        $ 2172 "Weight_value≔get_weight()" "noBreak"
        global Weight_value=get_weight()
        $ 2173 "tilt_angle≔-1" "noBreak"
        global tilt_angle=-1
        $ 2174 "Wait: 0.5" "noBreak"
        sleep(0.5)
        $ 2175 "vib_mot_thread≔ False " "noBreak"
        global vib_mot_thread=  False
        $ 2176 "MoveL" "noBreak"
        $ 2177 "dispense_pos" "noBreak"
        movel(dispense_pos, a=0.2, v=0.05)
        $ 2178 "Integral_error≔0" "noBreak"
        global Integral_error=0
        $ 2179 "current_error≔0" "noBreak"
        global current_error=0
        $ 2180 "previous_error≔0" "noBreak"
        global previous_error=0
        $ 2181 "Set AO[0]=0.0" "noBreak"
        set_standard_analog_out(0, 0.0)
        # begin: URCap Program Node
        #   Source: SensoPart VISOR Robotic, 2.0.0, SensoPart Industriesensorik GmbH
        #   Type: Exit Pose
        $ 2182 "Exit Pose" "noBreak"
        movel(pose_trans(easyPickPose,p[0.0000,0.0000,-0.0000,0.0000,0.0000,0.0000]),a=0.5000,v=0.2500,t=0.000000,r=0.000000)
        # end: URCap Program Node
        easyPickObjTaken = True
      end
      # end: URCap Program Node
      # begin: URCap Program Node
      #   Source: SensoPart VISOR Robotic, 2.0.0, SensoPart Industriesensorik GmbH
      #   Type: No Object Detected
      $ 2183 "No Object Detected" "noBreak"
      if (visor_partsFound(easyPickVisorId) < 1):
        $ 2184 "Popup: No weigh scale detected" "noBreak"
        popup("No weigh scale detected", "Message", False, False, blocking=True)
        else:
      end
      # end: URCap Program Node
    end
    easyPickCount_4 = easyPickCount_4 + 1
    visor_easyPickUpdate(easyPickVisorId, "counter", easyPickCount_4)
    visor_easyPickSetIdent("b1dffd", easyPickVisorId)
    # end: URCap Program Node
  end
  visorFuncEasyPick_a4e600()
  # end: URCap Program Node
  $ 2185 "powder dispensing"
  $ 2187 "Loop Weight_value<Target_weight"
  while (Weight_value<Target_weight):
    $ 2188 "MoveL"
    $ 2189 "Waypoint_75" "breakAfter"
    movel(Waypoint_75_p, a=0.3, v=0.05, r=0.05)
    $ 2190 "ftr_scoop2" "breakAfter"
    movel(ftr_scoop2_p, a=0.3, v=0.05)
    $ 2191 "aftr_scoop1" "breakAfter"
    movel(aftr_scoop1_p, a=0.3, v=0.05)
    $ 2192 "After_disp_3" "breakAfter"
    movel(After_disp_3_p, a=0.3, v=0.05)
    $ 2193 "Loop 1 times"
    Loop_13 = 0
    while (Loop_13 < 1):
      $ 2194 "Waypoint_55" "breakAfter"
      global move_thread_flag_2194=0
      thread move_thread_2194():
        enter_critical
        move_thread_flag_2194 = 1
        movel(Waypoint_55_p, a=0.5, v=0.07)
        move_thread_flag_2194 = 2
        exit_critical
      end
      move_thread_flag_2194 = 0
      move_thread_han_2194 = run move_thread_2194()
      while (True):
        sleep(1.0E-10)
        if (move_thread_flag_2194 > 1):
          join move_thread_han_2194
          break
        end
        sync()
      end
      $ 2196 "Waypoint_56" "breakAfter"
      movel(Waypoint_56_p, a=0.3, v=0.05)
      $ 2197 "Waypoint_74" "breakAfter"
      movel(Waypoint_74_p, a=0.3, v=0.05)
      $ 2198 "Set AO[0]=3.0"
      set_standard_analog_out(0, 0.3)
      $ 2199 "Wait: 2.0"
      sleep(2.0)
      $ 2200 "Set AO[0]=0.0"
      set_standard_analog_out(0, 0.0)
      Loop_13 = Loop_13 + 1
    end
    $ 2201 "ftr_scoop2" "breakAfter"
    movel(ftr_scoop2_p, a=0.3, v=0.05)
    $ 2202 "aftr_scoo3" "breakAfter"
    movel(aftr_scoo3_p, a=0.3, v=0.05)
    $ 2203 "MoveJ"
    $ 2204 "Waypoint_60" "breakAfter"
    movej(get_inverse_kin(Waypoint_60_p, qnear=Waypoint_60_q), a=0.5235987755982988, v=0.3490658503988659, r=0.05)
    $ 2205 "Waypoint_61" "breakAfter"
    movej(get_inverse_kin(Waypoint_61_p, qnear=Waypoint_61_q), a=0.5235987755982988, v=0.3490658503988659, r=0.05)
    $ 2206 "Waypoint_62" "breakAfter"
    movej(get_inverse_kin(Waypoint_62_p, qnear=Waypoint_62_q), a=0.5235987755982988, v=0.3490658503988659)
    $ 2207 "MoveL"
    $ 2208 "Start_thread≔ True "
    global Start_thread=  True
    $ 2209 "dispense_pos" "breakAfter"
    movel(dispense_pos, a=0.2, v=0.05)
    $ 2210 "vib_mot_thread≔ True "
    global vib_mot_thread=  True
    $ 2211 "Wait: 0.5"
    sleep(0.5)
    $ 2212 "Loop Weight_value≤Target_weight and tilt_angle≤-0.40"
    thread Thread_while_2212():
      while (True):
        $ 2213 "current_error≔Target_weight-Weight_value"
        global current_error=Target_weight-Weight_value
        $ 2214 "Integral_error≔Integral_error+current_error*dt"
        global Integral_error=Integral_error+current_error*dt
        $ 2215 "derivative≔(current_error-previous_error)/dt"
        global derivative=(current_error-previous_error)/dt
        $ 2216 "tilt_increment≔(kp*current_error)+(ki*Integral_error)+(kd*derivative)"
        global tilt_increment=(kp*current_error)+(ki*Integral_error)+(kd*derivative)
        $ 2217 "current_pose≔get_actual_tcp_pose()"
        global current_pose= get_actual_tcp_pose ()
        $ 2218 "tilt_angle≔current_pose[4]"
        global tilt_angle=current_pose[4]
        $ 2219 "tilt_pose≔pose_trans(current_pose, p[(tilt_increment/7), 0, 0, 0, tilt_increment, 0])"
        global tilt_pose=pose_trans(current_pose, p[(tilt_increment/7), 0, 0, 0, tilt_increment, 0])
        $ 2220 "movel(tilt_pose, a=0.025, v=0.015, r=0.00001)"
        movel(tilt_pose, a=0.025, v=0.015, r=0.00001)
        $ 2221 "previous_error≔current_error"
        global previous_error=current_error
        $ 2222 "Wait: 0.01"
        sleep(0.01)
      end
    end
    if (Weight_value <= Target_weight  and  tilt_angle <= -0.40):
      global thread_handler_2212=run Thread_while_2212()
      while (Weight_value <= Target_weight  and  tilt_angle <= -0.40):
        sync()
      end
      kill thread_handler_2212
    end
    $ 2223 "Start_thread≔ False "
    global Start_thread=  False
    $ 2224 "Set AO[0]=0.0"
    set_standard_analog_out(0, 0.0)
    $ 2225 "vib_mot_thread≔ False "
    global vib_mot_thread=  False
    $ 2227 "Weight_value≔get_weight()"
    global Weight_value=get_weight()
    $ 2228 "tilt_angle≔-1"
    global tilt_angle=-1
    $ 2229 "Wait: 0.5"
    sleep(0.5)
    $ 2230 "MoveL"
    $ 2231 "dispense_pos" "breakAfter"
    movel(dispense_pos, a=0.2, v=0.05)
    $ 2232 "Integral_error≔0"
    global Integral_error=0
    $ 2233 "current_error≔0"
    global current_error=0
    $ 2234 "previous_error≔0"
    global previous_error=0
  end
  $ 2235 "MoveL"
  $ 2236 "aftr_scoo3" "breakAfter"
  movel(aftr_scoo3_p, a=0.3, v=0.1)
  $ 2237 "ftr_scoop2" "breakAfter"
  movel(ftr_scoop2_p, a=0.4, v=0.1)
  $ 2238 "aftr_scoop1" "breakAfter"
  movel(aftr_scoop1_p, a=0.4, v=0.1)
  $ 2239 "After_disp_3" "breakAfter"
  movel(After_disp_3_p, a=0.4, v=0.1)
  $ 2240 "Set AO[0]=3.0"
  set_standard_analog_out(0, 0.3)
  $ 2241 "Wait: 2.0"
  sleep(2.0)
  $ 2242 "Set AO[0]=0.0"
  set_standard_analog_out(0, 0.0)
  $ 2243 "aftr_scoop1" "breakAfter"
  movel(aftr_scoop1_p, a=1.2, v=0.25)
  $ 2244 "ftr_scoop2" "breakAfter"
  movel(ftr_scoop2_p, a=0.4, v=0.1)
  $ 2245 "Waypoint_63" "breakAfter"
  movel(Waypoint_63_p, a=1.2, v=0.25, r=0.05)
  $ 2246 "Start" "breakAfter"
  movel(Start_p, a=0.6, v=0.15)
  $ 2247 "Popup: Powder dispensed successfully..."
  popup("Powder dispensed successfully...", "Message", False, False, blocking=True)
  elif (38 == switch_1):
    $ 2248 "Case 38"
    $ 2249 "PowderA(M200)"
    # begin: URCap Program Node
    #   Source: SensoPart VISOR Robotic, 2.0.0, SensoPart Industriesensorik GmbH
    #   Type: VISOR Robotic App
    $ 2250 "VISOR Easy Pick"
    def visorFuncEasyPick_cfdeea():
      # begin: URCap Program Node
      #   Source: SensoPart VISOR Robotic, 2.0.0, SensoPart Industriesensorik GmbH
      #   Type: Easy Pick Setup
      $ 2251 "# 1 Setup" "noBreak"
      local easyPickVisorId = 1
      local easyPickArmMounted = True
      local easyPickSetJob = True
      local easyPickJobName = "PowderA"
      local easyPickAtImgAcq = False
      local easyPickImgAcqPose = cont_img_pose
      # end: URCap Program Node
      # begin: URCap Program Node
      #   Source: SensoPart VISOR Robotic, 2.0.0, SensoPart Industriesensorik GmbH
      #   Type: Process
      $ 2252 "Process" "noBreak"
      local easyPickObjTaken = False
      local easyPickTrigger = False
      local easyPickPoseIdx = 0
      local easyPickPose = p[0,0,0,0,0,0]
      def easyPickFuncTrigger(visorId, setJob, jobName, arm):
      if (setJob):
        visor_changeJob(visorId, jobName, 6000)
      end
      if (arm):
        visor_trigger(visorId, 6000, "arm")
      else:
        visor_trigger(visorId, 6000)
      end
      global easyPickParts_6=visor_partsFound(visorId)
      visor_easyPickUpdate(visorId, "parts", visor_partsFound(visorId))
      return visor_getPose3d(visorId, 0)
    end
    while (not easyPickObjTaken):
      easyPickTrigger = (easyPickCount_6 >= visor_partsFound(easyPickVisorId)) or (easyPickCount_6 > 9) or (not visor_easyPickCheckIdent("9c10c0", easyPickVisorId))
      if (easyPickTrigger):
        easyPickCount_6 = 0
      end
      easyPickPoseIdx = easyPickCount_6
      easyPickPose = visor_getPose3d(easyPickVisorId, easyPickPoseIdx)
      visor_easyPickUpdate(easyPickVisorId, "counter", easyPickPoseIdx)
      # begin: URCap Program Node
      #   Source: SensoPart VISOR Robotic, 2.0.0, SensoPart Industriesensorik GmbH
      #   Type: Image Acquisition Pose
      $ 2253 "Image Acquisition Pose" "noBreak"
      if (easyPickTrigger):
        if (not easyPickAtImgAcq):
          movej(pose_trans(easyPickImgAcqPose,p[0.0000,0.0000,-0.0000,0.0000,0.0000,0.0000]),a=1.3963,v=1.0472,t=0.000000,r=0.000000)
          easyPickAtImgAcq = True
        end
        easyPickPose = easyPickFuncTrigger(easyPickVisorId, easyPickSetJob, easyPickJobName, easyPickArmMounted)
      end
      # end: URCap Program Node
      # begin: URCap Program Node
      #   Source: SensoPart VISOR Robotic, 2.0.0, SensoPart Industriesensorik GmbH
      #   Type: Object Detected
      $ 2254 "Object Detected" "noBreak"
      if (visor_partsFound(easyPickVisorId) > 0):
        $ 2255 "Open Gripper" "noBreak"
        # begin: URCap Program Node
        #   Source: Robotiq_Grippers, 1.8.4.4844, Robotiq Inc.
        #   Type: Gripper
        $ 2256 "Gripper Open (1)" "noBreak"
        if not(gripper_connected[0]):
          popup("Gripper 1 must be connected to run this program.", "No connection", False, True, True)
        end
        if not(rq_is_gripper_activated("1")):
          popup("Gripper 1 is not activated. Go to Installation tab > Gripper to activate it and run the program again.", "Not activated", False, True, True)
        end
        rq_set_pos_spd_for(0, 77, 77, "1")
        rq_wait_pos_spe_for_request(0, 77, 77, "1")
        rq_go_to("1")
        rq_wait("1")
        # end: URCap Program Node
        $ 2257 "MoveJ" "noBreak"
        $ 2258 "Waypoint_76" "noBreak"
        movej(get_inverse_kin(Waypoint_76_p, qnear=Waypoint_76_q), a=1.3962634015954636, v=1.0471975511965976)
        # begin: URCap Program Node
        #   Source: SensoPart VISOR Robotic, 2.0.0, SensoPart Industriesensorik GmbH
        #   Type: Approach Pose
        $ 2259 "Approach Pose" "noBreak"
        movej(pose_trans(easyPickPose,p[0.0000,0.0000,0.0500,0.0000,0.0000,0.0000]),a=1.3963,v=1.0472,t=0.000000,r=0.000000)
        # end: URCap Program Node
        # begin: URCap Program Node
        #   Source: SensoPart VISOR Robotic, 2.0.0, SensoPart Industriesensorik GmbH
        #   Type: Target Pose
        $ 2260 "Target Pose" "noBreak"
        movel(pose_trans(easyPickPose,p[0.0000,0.0000,-0.0000,0.0000,0.0000,0.0000]),a=0.5000,v=0.2500,t=0.000000,r=0.000000)
        # end: URCap Program Node
        $ 2261 "Close Gripper" "noBreak"
        # begin: URCap Program Node
        #   Source: Robotiq_Grippers, 1.8.4.4844, Robotiq Inc.
        #   Type: Gripper
        $ 2262 "Gripper Move0mm (1)" "noBreak"
        if not(gripper_connected[0]):
          popup("Gripper 1 must be connected to run this program.", "No connection", False, True, True)
        end
        if not(rq_is_gripper_activated("1")):
          popup("Gripper 1 is not activated. Go to Installation tab > Gripper to activate it and run the program again.", "Not activated", False, True, True)
        end
        rq_set_pos_spd_for(247, 77, 77, "1")
        rq_wait_pos_spe_for_request(247, 77, 77, "1")
        rq_go_to("1")
        rq_wait("1")
        # end: URCap Program Node
        # begin: URCap Program Node
        #   Source: SensoPart VISOR Robotic, 2.0.0, SensoPart Industriesensorik GmbH
        #   Type: Exit Pose
        $ 2263 "Exit Pose" "noBreak"
        movel(pose_trans(easyPickPose,p[0.0000,0.0000,0.0500,0.0000,0.0000,0.0000]),a=0.5000,v=0.2500,t=0.000000,r=0.000000)
        # end: URCap Program Node
        easyPickObjTaken = True
      end
      # end: URCap Program Node
      # begin: URCap Program Node
      #   Source: SensoPart VISOR Robotic, 2.0.0, SensoPart Industriesensorik GmbH
      #   Type: No Object Detected
      $ 2264 "No Object Detected" "noBreak"
      if (visor_partsFound(easyPickVisorId) < 1):
        $ 2265 "Popup: No Powder container is detected" "noBreak"
        popup("No Powder container is detected", "Message", False, False, blocking=True)
        else:
      end
      # end: URCap Program Node
    end
    easyPickCount_6 = easyPickCount_6 + 1
    visor_easyPickUpdate(easyPickVisorId, "counter", easyPickCount_6)
    visor_easyPickSetIdent("9c10c0", easyPickVisorId)
    # end: URCap Program Node
  end
  visorFuncEasyPick_cfdeea()
  # end: URCap Program Node
  $ 2266 "MoveJ"
  $ 2267 "PowderA_wayp1" "breakAfter"
  movej(get_inverse_kin(PowderA_wayp1_p, qnear=PowderA_wayp1_q), a=1.3962634015954636, v=1.0471975511965976, r=0.05)
  $ 2268 "MoveL"
  $ 2269 "Waypoint_80" "breakAfter"
  movel(Waypoint_80_p, a=1.2, v=0.25)
  $ 2270 "MoveL"
  $ 2271 "Decapp_above" "breakAfter"
  movel(Decapp_above_p, a=1.2, v=0.25)
  $ 2272 "Set GRP_3F_Open=On"
  set_standard_digital_out(5, True)
  $ 2273 "Wait: 0.5"
  sleep(0.5)
  $ 2274 "Decapp_place" "breakAfter"
  movel(Decapp_place_p, a=0.3, v=0.05)
  $ 2275 "Set GRP_3F_Open=Off"
  set_standard_digital_out(5, False)
  $ 2276 "Wait: 0.5"
  sleep(0.5)
  # begin: URCap Program Node
  #   Source: Robotiq_Grippers, 1.8.4.4844, Robotiq Inc.
  #   Type: Gripper
  $ 2277 "Gripper Move40mm (1)"
  if not(gripper_connected[0]):
    popup("Gripper 1 must be connected to run this program.", "No connection", False, True, True)
  end
  if not(rq_is_gripper_activated("1")):
    popup("Gripper 1 is not activated. Go to Installation tab > Gripper to activate it and run the program again.", "Not activated", False, True, True)
  end
  rq_set_pos_spd_for(64, 77, 77, "1")
  rq_wait_pos_spe_for_request(64, 77, 77, "1")
  rq_go_to("1")
  rq_wait("1")
  # end: URCap Program Node
  $ 2278 "MoveL"
  $ 2279 "Decapp_above" "breakAfter"
  movel(Decapp_above_p, a=1.2, v=0.25)
  $ 2280 "Waypoint_78" "breakAfter"
  movel(Waypoint_78_p, a=1.2, v=0.25, r=0.05)
  $ 2281 "Home (Safe)"
  movej([-1.2302089344500047, -1.2969853503591224, -1.875639182904262, -1.539621866126728, 1.5731943360401213, -2.80099559440227], a=1.3962634015954636, v=1.0471975511965976)
  elif (39 == switch_1):
    $ 2282 "Case 39"
    $ 2283 "Decap Container A"
    $ 2284 "MoveL"
    $ 2285 "Waypoint_81" "breakAfter"
    movel(Waypoint_81_p, a=1.2, v=0.25)
    $ 2286 "Waypoint_79" "breakAfter"
    movel(Waypoint_79_p, a=1.2, v=0.25)
    # begin: URCap Program Node
    #   Source: Robotiq_Grippers, 1.8.4.4844, Robotiq Inc.
    #   Type: Gripper
    $ 2287 "Gripper Move22mm (1)"
    if not(gripper_connected[0]):
      popup("Gripper 1 must be connected to run this program.", "No connection", False, True, True)
    end
    if not(rq_is_gripper_activated("1")):
      popup("Gripper 1 is not activated. Go to Installation tab > Gripper to activate it and run the program again.", "Not activated", False, True, True)
    end
    rq_set_pos_spd_for(145, 77, 77, "1")
    rq_wait_pos_spe_for_request(145, 77, 77, "1")
    rq_go_to("1")
    rq_wait("1")
    # end: URCap Program Node
    $ 2288 "Decap"
    $ 2289 "Action_Info≔'decapping'"
    global Action_Info="decapping"
    $ 2290 "Set GRP_3F_Enable=On"
    set_standard_digital_out(4, True)
    $ 2291 "Set GRP_3F_Decap=On"
    set_standard_digital_out(3, True)
    $ 2292 "Force"
    sleep(0.02)
    zero_ftsensor()
    force_mode(p[0.0,0.0,0.0,0.0,0.0,0.0], [0, 0, 1, 0, 0, 0], [0.0, 0.0, 2.0, 0.0, 0.0, 0.0], 2, [0.1, 0.1, 5.0E-4, 0.3490658503988659, 0.3490658503988659, 0.3490658503988659])
    $ 2293 "check_decapping(offset=0.010, timeout=4, abort=CMD_Hold)" "noBreak"
    check_decapping(offset=0.010, timeout=4, abort=CMD_Hold)
    end_force_mode()
    stopl(5.0)
    $ 2294 "Set GRP_3F_Decap=Off"
    set_standard_digital_out(3, False)
    $ 2295 "Set GRP_3F_Enable=Off"
    set_standard_digital_out(4, False)
    $ 2296 "MoveL"
    $ 2297 "Waypoint_82" "breakAfter"
    movel(Waypoint_82_p, a=1.2, v=0.25)
    $ 2298 "Cap_above" "breakAfter"
    movel(Cap_above_p, a=1.2, v=0.25, r=0.05)
    $ 2299 "Cap_Place" "breakAfter"
    movel(Cap_Place_p, a=1.2, v=0.25)
    # begin: URCap Program Node
    #   Source: Robotiq_Grippers, 1.8.4.4844, Robotiq Inc.
    #   Type: Gripper
    $ 2300 "Gripper Move39mm (1)"
    if not(gripper_connected[0]):
      popup("Gripper 1 must be connected to run this program.", "No connection", False, True, True)
    end
    if not(rq_is_gripper_activated("1")):
      popup("Gripper 1 is not activated. Go to Installation tab > Gripper to activate it and run the program again.", "Not activated", False, True, True)
    end
    rq_set_pos_spd_for(67, 77, 77, "1")
    rq_wait_pos_spe_for_request(67, 77, 77, "1")
    rq_go_to("1")
    rq_wait("1")
    # end: URCap Program Node
    $ 2301 "Cap_above" "breakAfter"
    movel(Cap_above_p, a=1.2, v=0.25)
    $ 2302 "Home (Safe)"
    movej([-1.2302089344500047, -1.2969853503591224, -1.875639182904262, -1.539621866126728, 1.5731943360401213, -2.80099559440227], a=1.3962634015954636, v=1.0471975511965976)
  elif (40 == switch_1):
    $ 2338 "Case 40"
    $ 2339 "Place the open PowderA container & dosing"
    # begin: URCap Program Node
    #   Source: SensoPart VISOR Robotic, 2.0.0, SensoPart Industriesensorik GmbH
    #   Type: VISOR Robotic App
    $ 2342 "VISOR Easy Pick"
    def visorFuncEasyPick_303fc5():
      # begin: URCap Program Node
      #   Source: SensoPart VISOR Robotic, 2.0.0, SensoPart Industriesensorik GmbH
      #   Type: Easy Pick Setup
      $ 2343 "# 1 Setup" "noBreak"
      local easyPickVisorId = 1
      local easyPickArmMounted = True
      local easyPickSetJob = True
      local easyPickJobName = "PoTS"
      local easyPickAtImgAcq = False
      local easyPickImgAcqPose = cont_img_pose
      # end: URCap Program Node
      # begin: URCap Program Node
      #   Source: SensoPart VISOR Robotic, 2.0.0, SensoPart Industriesensorik GmbH
      #   Type: Process
      $ 2344 "Process" "noBreak"
      local easyPickObjTaken = False
      local easyPickTrigger = False
      local easyPickPoseIdx = 0
      local easyPickPose = p[0,0,0,0,0,0]
      def easyPickFuncTrigger(visorId, setJob, jobName, arm):
      if (setJob):
        visor_changeJob(visorId, jobName, 6000)
      end
      if (arm):
        visor_trigger(visorId, 6000, "arm")
      else:
        visor_trigger(visorId, 6000)
      end
      global easyPickParts_7=visor_partsFound(visorId)
      visor_easyPickUpdate(visorId, "parts", visor_partsFound(visorId))
      return visor_getPose3d(visorId, 0)
    end
    while (not easyPickObjTaken):
      easyPickTrigger = (easyPickCount_7 >= visor_partsFound(easyPickVisorId)) or (easyPickCount_7 > 9) or (not visor_easyPickCheckIdent("2f5077", easyPickVisorId))
      if (easyPickTrigger):
        easyPickCount_7 = 0
      end
      easyPickPoseIdx = easyPickCount_7
      easyPickPose = visor_getPose3d(easyPickVisorId, easyPickPoseIdx)
      visor_easyPickUpdate(easyPickVisorId, "counter", easyPickPoseIdx)
      # begin: URCap Program Node
      #   Source: SensoPart VISOR Robotic, 2.0.0, SensoPart Industriesensorik GmbH
      #   Type: Image Acquisition Pose
      $ 2345 "Image Acquisition Pose" "noBreak"
      if (easyPickTrigger):
        if (not easyPickAtImgAcq):
          movej(pose_trans(easyPickImgAcqPose,p[0.0000,0.0000,-0.0000,0.0000,0.0000,0.0000]),a=1.3963,v=1.0472,t=0.000000,r=0.000000)
          easyPickAtImgAcq = True
        end
        easyPickPose = easyPickFuncTrigger(easyPickVisorId, easyPickSetJob, easyPickJobName, easyPickArmMounted)
      end
      # end: URCap Program Node
      # begin: URCap Program Node
      #   Source: SensoPart VISOR Robotic, 2.0.0, SensoPart Industriesensorik GmbH
      #   Type: Object Detected
      $ 2346 "Object Detected" "noBreak"
      if (visor_partsFound(easyPickVisorId) > 0):
        $ 2347 "Open Gripper" "noBreak"
        # begin: URCap Program Node
        #   Source: Robotiq_Grippers, 1.8.4.4844, Robotiq Inc.
        #   Type: Gripper
        $ 2348 "Gripper Open (1)" "noBreak"
        if not(gripper_connected[0]):
          popup("Gripper 1 must be connected to run this program.", "No connection", False, True, True)
        end
        if not(rq_is_gripper_activated("1")):
          popup("Gripper 1 is not activated. Go to Installation tab > Gripper to activate it and run the program again.", "Not activated", False, True, True)
        end
        rq_set_pos_spd_for(0, 77, 77, "1")
        rq_wait_pos_spe_for_request(0, 77, 77, "1")
        rq_go_to("1")
        rq_wait("1")
        # end: URCap Program Node
        $ 2349 "MoveL" "noBreak"
        $ 2350 "OP_PowderA2" "noBreak"
        movel(OP_PowderA2_p, a=1.2, v=0.25)
        $ 2351 "OP_PowderA_abov" "noBreak"
        movel(OP_PowderA_abov_p, a=1.2, v=0.25)
        $ 2352 "OP_PowderA_pick" "noBreak"
        movel(OP_PowderA_pick_p, a=1.2, v=0.25)
        # begin: URCap Program Node
        #   Source: Robotiq_Grippers, 1.8.4.4844, Robotiq Inc.
        #   Type: Gripper
        $ 2353 "Gripper Close (1)" "noBreak"
        if not(gripper_connected[0]):
          popup("Gripper 1 must be connected to run this program.", "No connection", False, True, True)
        end
        if not(rq_is_gripper_activated("1")):
          popup("Gripper 1 is not activated. Go to Installation tab > Gripper to activate it and run the program again.", "Not activated", False, True, True)
        end
        rq_set_pos_spd_for(255, 77, 77, "1")
        rq_wait_pos_spe_for_request(255, 77, 77, "1")
        rq_go_to("1")
        rq_wait("1")
        # end: URCap Program Node
        $ 2354 "Wait: 0.5" "noBreak"
        sleep(0.5)
        $ 2355 "Set GRP_3F_Open=On" "noBreak"
        set_standard_digital_out(5, True)
        $ 2357 "OP_PowderA_abov" "noBreak"
        movel(OP_PowderA_abov_p, a=0.3, v=0.05)
        $ 2358 "Op_PowA_wP" "noBreak"
        movel(Op_PowA_wP_p, a=1.2, v=0.25)
        # begin: URCap Program Node
        #   Source: SensoPart VISOR Robotic, 2.0.0, SensoPart Industriesensorik GmbH
        #   Type: Approach Pose
        $ 2359 "Approach Pose" "noBreak"
        movej(pose_trans(easyPickPose,p[0.0000,0.0000,-0.0000,0.0000,0.0000,0.0000]),a=0.5236,v=0.4363,t=0.000000,r=0.000000)
        # end: URCap Program Node
        # begin: URCap Program Node
        #   Source: SensoPart VISOR Robotic, 2.0.0, SensoPart Industriesensorik GmbH
        #   Type: Target Pose
        $ 2360 "Target Pose" "noBreak"
        movel(pose_trans(easyPickPose,p[0.0000,0.0000,-0.0000,0.0000,0.0000,0.0000]),a=0.1000,v=0.0500,t=0.000000,r=0.000000)
        # end: URCap Program Node
        $ 2361 "Close Gripper" "noBreak"
        $ 2362 "target_pose≔pose_add(get_actual_tcp_pose(), p[0,0,-0.085,0,0,0])" "noBreak"
        global target_pose=pose_add(get_actual_tcp_pose(), p[0,0,-0.085,0,0,0])
        $ 2363 "MoveL" "noBreak"
        $ 2364 "target_pose" "noBreak"
        movel(target_pose, a=0.3, v=0.05)
        # begin: URCap Program Node
        #   Source: Robotiq_Grippers, 1.8.4.4844, Robotiq Inc.
        #   Type: Gripper
        $ 2365 "Gripper Open (1)" "noBreak"
        if not(gripper_connected[0]):
          popup("Gripper 1 must be connected to run this program.", "No connection", False, True, True)
        end
        if not(rq_is_gripper_activated("1")):
          popup("Gripper 1 is not activated. Go to Installation tab > Gripper to activate it and run the program again.", "Not activated", False, True, True)
        end
        rq_set_pos_spd_for(0, 77, 77, "1")
        rq_wait_pos_spe_for_request(0, 77, 77, "1")
        rq_go_to("1")
        rq_wait("1")
        # end: URCap Program Node
        # begin: URCap Program Node
        #   Source: SensoPart VISOR Robotic, 2.0.0, SensoPart Industriesensorik GmbH
        #   Type: Exit Pose
        $ 2366 "Exit Pose" "noBreak"
        movel(pose_trans(easyPickPose,p[0.0000,0.0000,-0.0000,0.0000,0.0000,0.0000]),a=0.5000,v=0.2500,t=0.000000,r=0.000000)
        # end: URCap Program Node
        easyPickObjTaken = True
      end
      # end: URCap Program Node
      # begin: URCap Program Node
      #   Source: SensoPart VISOR Robotic, 2.0.0, SensoPart Industriesensorik GmbH
      #   Type: No Object Detected
      $ 2367 "No Object Detected" "noBreak"
      if (visor_partsFound(easyPickVisorId) < 1):
        $ 2368 "Popup: No weigh scale detected" "noBreak"
        popup("No weigh scale detected", "Message", False, False, blocking=True)
        else:
      end
      # end: URCap Program Node
    end
    easyPickCount_7 = easyPickCount_7 + 1
    visor_easyPickUpdate(easyPickVisorId, "counter", easyPickCount_7)
    visor_easyPickSetIdent("2f5077", easyPickVisorId)
    # end: URCap Program Node
  end
  visorFuncEasyPick_303fc5()
  # end: URCap Program Node
  $ 2369 "place_pose≔get_actual_tcp_pose()"
  global place_pose= get_actual_tcp_pose ()
  $ 2370 "center_pose()"
  center_pose()
  $ 2371 "center_pose_t≔P_center"
  global center_pose_t=P_center
  $ 2372 "MoveJ"
  $ 2373 "Waypoint_1" "breakAfter"
  movej(get_inverse_kin(Waypoint_1_p, qnear=Waypoint_1_q), a=1.3962634015954636, v=1.0471975511965976)
  elif (41 == switch_1):
    $ 2374 "Case 41"
    $ 2375 "Powder Emptying"
    $ 2376 "zero_scale()"
    zero_scale()
    $ 2377 "Task≔'Emptying'"
    global Task="Emptying"
    # begin: URCap Program Node
    #   Source: SensoPart VISOR Robotic, 2.0.0, SensoPart Industriesensorik GmbH
    #   Type: VISOR Robotic App
    $ 2378 "VISOR Easy Pick"
    def visorFuncEasyPick_221058():
      # begin: URCap Program Node
      #   Source: SensoPart VISOR Robotic, 2.0.0, SensoPart Industriesensorik GmbH
      #   Type: Easy Pick Setup
      $ 2379 "# 1 Setup" "noBreak"
      local easyPickVisorId = 1
      local easyPickArmMounted = True
      local easyPickSetJob = True
      local easyPickJobName = "Weigh_target"
      local easyPickAtImgAcq = False
      local easyPickImgAcqPose = FRM_Weigh_scale
      # end: URCap Program Node
      # begin: URCap Program Node
      #   Source: SensoPart VISOR Robotic, 2.0.0, SensoPart Industriesensorik GmbH
      #   Type: Process
      $ 2380 "Process" "noBreak"
      local easyPickObjTaken = False
      local easyPickTrigger = False
      local easyPickPoseIdx = 0
      local easyPickPose = p[0,0,0,0,0,0]
      def easyPickFuncTrigger(visorId, setJob, jobName, arm):
      if (setJob):
        visor_changeJob(visorId, jobName, 6000)
      end
      if (arm):
        visor_trigger(visorId, 6000, "arm")
      else:
        visor_trigger(visorId, 6000)
      end
      global easyPickParts_4=visor_partsFound(visorId)
      visor_easyPickUpdate(visorId, "parts", visor_partsFound(visorId))
      return visor_getPose3d(visorId, 0)
    end
    while (not easyPickObjTaken):
      easyPickTrigger = (easyPickCount_4 >= visor_partsFound(easyPickVisorId)) or (easyPickCount_4 > 9) or (not visor_easyPickCheckIdent("7aa8bf", easyPickVisorId))
      if (easyPickTrigger):
        easyPickCount_4 = 0
      end
      easyPickPoseIdx = easyPickCount_4
      easyPickPose = visor_getPose3d(easyPickVisorId, easyPickPoseIdx)
      visor_easyPickUpdate(easyPickVisorId, "counter", easyPickPoseIdx)
      # begin: URCap Program Node
      #   Source: SensoPart VISOR Robotic, 2.0.0, SensoPart Industriesensorik GmbH
      #   Type: Image Acquisition Pose
      $ 2381 "Image Acquisition Pose" "noBreak"
      if (easyPickTrigger):
        if (not easyPickAtImgAcq):
          movej(pose_trans(easyPickImgAcqPose,p[0.0000,0.0000,-0.0000,0.0000,0.0000,0.0000]),a=1.3963,v=1.0472,t=0.000000,r=0.000000)
          easyPickAtImgAcq = True
        end
        easyPickPose = easyPickFuncTrigger(easyPickVisorId, easyPickSetJob, easyPickJobName, easyPickArmMounted)
      end
      # end: URCap Program Node
      # begin: URCap Program Node
      #   Source: SensoPart VISOR Robotic, 2.0.0, SensoPart Industriesensorik GmbH
      #   Type: Object Detected
      $ 2382 "Object Detected" "noBreak"
      if (visor_partsFound(easyPickVisorId) > 0):
        $ 2383 "Open Gripper" "noBreak"
        $ 2384 "tare_scale()" "noBreak"
        tare_scale()
        $ 2385 "Wait: 0.2" "noBreak"
        sleep(0.2)
        $ 2386 "Weight_value≔get_weight()" "noBreak"
        global Weight_value=get_weight()
        $ 2387 "Wait: 0.2" "noBreak"
        sleep(0.2)
        $ 2388 "compute_level_percent(W_now, Weight_value)" "noBreak"
        compute_level_percent(W_now, Weight_value)
        $ 2389 "If level≥10.0" "noBreak"
        if (level >= 10.0):
          $ 2390 "MoveJ" "noBreak"
          $ 2391 "Spatula_otw" "noBreak"
          movej(get_inverse_kin(Spatula_otw_p, qnear=Spatula_otw_q), a=1.3962634015954636, v=1.0471975511965976)
          $ 2392 "pick_spat_L_abv" "noBreak"
          movej(get_inverse_kin(pick_spat_L_abv_p, qnear=pick_spat_L_abv_q), a=1.3962634015954636, v=1.0471975511965976)
          $ 2393 "MoveL" "noBreak"
          $ 2394 "spat_L_pick" "noBreak"
          movel(spat_L_pick_p, a=1.2, v=0.25)
          # begin: URCap Program Node
          #   Source: Robotiq_Grippers, 1.8.4.4844, Robotiq Inc.
          #   Type: Gripper
          $ 2395 "Gripper Close (1)" "noBreak"
          if not(gripper_connected[0]):
            popup("Gripper 1 must be connected to run this program.", "No connection", False, True, True)
          end
          if not(rq_is_gripper_activated("1")):
            popup("Gripper 1 is not activated. Go to Installation tab > Gripper to activate it and run the program again.", "Not activated", False, True, True)
          end
          rq_set_pos_spd_for(255, 0, 77, "1")
          rq_wait_pos_spe_for_request(255, 0, 77, "1")
          rq_go_to("1")
          rq_wait("1")
          # end: URCap Program Node
          $ 2396 "spat_L_lift" "noBreak"
          movel(spat_L_lift_p, a=1.2, v=0.25)
          $ 2397 "spat_L_side" "noBreak"
          movel(spat_L_side_p, a=1.2, v=0.25)
          $ 2398 "spat_L_up" "noBreak"
          movel(spat_L_up_p, a=1.2, v=0.25)
          $ 2399 "MoveJ" "noBreak"
          $ 2400 "Spatula_otw" "noBreak"
          movej(get_inverse_kin(Spatula_otw_p, qnear=Spatula_otw_q), a=1.3962634015954636, v=1.0471975511965976)
        else:
          $ 2401 "ElseIf level≥1.0  and level<10.0" "noBreak"
          if (level >= 1.0   and  level<10.0):
            $ 2402 "MoveJ" "noBreak"
            $ 2403 "Spatula_otw" "noBreak"
            movej(get_inverse_kin(Spatula_otw_p, qnear=Spatula_otw_q), a=1.3962634015954636, v=1.0471975511965976)
            $ 2404 "spat_M_up" "noBreak"
            movej(get_inverse_kin(spat_M_up_p, qnear=spat_M_up_q), a=1.3962634015954636, v=1.0471975511965976)
            $ 2405 "MoveL" "noBreak"
            $ 2406 "spat_M_pick" "noBreak"
            movel(spat_M_pick_p, a=1.2, v=0.25)
            # begin: URCap Program Node
            #   Source: Robotiq_Grippers, 1.8.4.4844, Robotiq Inc.
            #   Type: Gripper
            $ 2407 "Gripper Close (1)" "noBreak"
            if not(gripper_connected[0]):
              popup("Gripper 1 must be connected to run this program.", "No connection", False, True, True)
            end
            if not(rq_is_gripper_activated("1")):
              popup("Gripper 1 is not activated. Go to Installation tab > Gripper to activate it and run the program again.", "Not activated", False, True, True)
            end
            rq_set_pos_spd_for(255, 0, 77, "1")
            rq_wait_pos_spe_for_request(255, 0, 77, "1")
            rq_go_to("1")
            rq_wait("1")
            # end: URCap Program Node
            $ 2408 "spat_M_up" "noBreak"
            movel(spat_M_up_p, a=1.2, v=0.25)
            $ 2409 "Spatula_otw" "noBreak"
            movel(Spatula_otw_p, a=1.2, v=0.25)
            $ 2410 "switch_spat_M≔ False " "noBreak"
            global switch_spat_M=  False
          else:
            $ 2411 "Else" "noBreak"
            $ 2412 "MoveJ" "noBreak"
            $ 2413 "Spatula_otw" "noBreak"
            movej(get_inverse_kin(Spatula_otw_p, qnear=Spatula_otw_q), a=1.3962634015954636, v=1.0471975511965976)
            $ 2414 "spat_S_up" "noBreak"
            movej(get_inverse_kin(spat_S_up_p, qnear=spat_S_up_q), a=1.3962634015954636, v=1.0471975511965976)
            $ 2415 "MoveL" "noBreak"
            $ 2416 "spat_S_pick" "noBreak"
            movel(spat_S_pick_p, a=1.2, v=0.25)
            # begin: URCap Program Node
            #   Source: Robotiq_Grippers, 1.8.4.4844, Robotiq Inc.
            #   Type: Gripper
            $ 2417 "Gripper Close (1)" "noBreak"
            if not(gripper_connected[0]):
              popup("Gripper 1 must be connected to run this program.", "No connection", False, True, True)
            end
            if not(rq_is_gripper_activated("1")):
              popup("Gripper 1 is not activated. Go to Installation tab > Gripper to activate it and run the program again.", "Not activated", False, True, True)
            end
            rq_set_pos_spd_for(255, 0, 77, "1")
            rq_wait_pos_spe_for_request(255, 0, 77, "1")
            rq_go_to("1")
            rq_wait("1")
            # end: URCap Program Node
            $ 2418 "spat_S_up" "noBreak"
            movel(spat_S_up_p, a=1.2, v=0.25)
            $ 2419 "Spatula_otw" "noBreak"
            movel(Spatula_otw_p, a=1.2, v=0.25)
            $ 2420 "switch_spat_S≔ False " "noBreak"
            global switch_spat_S=  False
          end
        end
        $ 2421 "Weight_value≔get_weight()" "noBreak"
        global Weight_value=get_weight()
        $ 2422 "auto_tilt_and_scoop(W_now, Target_weight, Weight_value)" "noBreak"
        auto_tilt_and_scoop(W_now, Target_weight, Weight_value)
        # begin: URCap Program Node
        #   Source: SensoPart VISOR Robotic, 2.0.0, SensoPart Industriesensorik GmbH
        #   Type: Approach Pose
        $ 2423 "Approach Pose" "noBreak"
        movej(pose_trans(easyPickPose,p[0.0000,0.0000,0.0500,0.0000,0.0000,0.0000]),a=0.2618,v=0.1745,t=0.000000,r=0.000000)
        # end: URCap Program Node
        # begin: URCap Program Node
        #   Source: SensoPart VISOR Robotic, 2.0.0, SensoPart Industriesensorik GmbH
        #   Type: Target Pose
        $ 2424 "Target Pose" "noBreak"
        movel(pose_trans(easyPickPose,p[0.0000,0.0000,-0.0000,0.0000,0.0000,0.0000]),a=0.0500,v=0.0200,t=0.000000,r=0.000000)
        # end: URCap Program Node
        $ 2425 "Close Gripper" "noBreak"
        $ 2426 "dispense_pos≔get_actual_tcp_pose()" "noBreak"
        global dispense_pos= get_actual_tcp_pose ()
        $ 2427 "Loop Weight_value≤Target_weight" "noBreak"
        while (Weight_value <= Target_weight):
          $ 2428 "MoveL" "noBreak"
          $ 2429 "dispense_pos" "noBreak"
          movel(dispense_pos, a=0.2, v=0.1)
          $ 2430 "log_weight()" "noBreak"
          log_weight()
          $ 2431 "Wait: 0.5" "noBreak"
          sleep(0.5)
          $ 2432 "If level≥90.0" "noBreak"
          if (level >= 90.0):
            $ 2433 "Rotate()" "noBreak"
            Rotate()
          end
          $ 2434 "If level≤70" "noBreak"
          if (level <= 70):
            $ 2435 "tilt_to_home()" "noBreak"
            tilt_to_home()
          end
          $ 2436 "Wait: 0.5" "noBreak"
          sleep(0.5)
          $ 2437 "Start_thread≔ True " "noBreak"
          global Start_thread=  True
          $ 2438 "vib_mot_thread≔ True " "noBreak"
          global vib_mot_thread=  True
          $ 2440 "Wait: 0.5" "noBreak"
          sleep(0.5)
          $ 2446 "If diff>0" "noBreak"
          if (diff>0):
            $ 2447 "tilt_pose≔pose_trans(get_actual_tcp_pose(), p[0, 0, 0, 0, 0, 2.0])" "noBreak"
            global tilt_pose=pose_trans(get_actual_tcp_pose(), p[0, 0, 0, 0, 0, 2.0])
            $ 2448 "movel(tilt_pose, a=0.1, v=0.1, r=0.00001)" "noBreak"
            movel(tilt_pose, a=0.1, v=0.1, r=0.00001)
          end
          $ 2460 "Start_thread≔ False " "noBreak"
          global Start_thread=  False
          $ 2462 "Weight_value≔get_weight()" "noBreak"
          global Weight_value=get_weight()
          $ 2464 "Wait: 0.5" "noBreak"
          sleep(0.5)
          $ 2465 "vib_mot_thread≔ False " "noBreak"
          global vib_mot_thread=  False
          $ 2466 "MoveL" "noBreak"
          $ 2467 "dispense_pos" "noBreak"
          movel(dispense_pos, a=0.5, v=0.25)
          $ 2468 "Integral_error≔0" "noBreak"
          global Integral_error=0
          $ 2469 "current_error≔0" "noBreak"
          global current_error=0
          $ 2470 "previous_error≔0" "noBreak"
          global previous_error=0
          $ 2471 "Set AO[0]=0.0" "noBreak"
          set_standard_analog_out(0, 0.0)
          $ 2472 "compute_level_percent(W_now, Weight_value)" "noBreak"
          compute_level_percent(W_now, Weight_value)
          $ 2473 "If spatula ≟ 'spatula_M'  and switch_spat_M≟ True " "noBreak"
          if (spatula  ==  "spatula_M"   and  switch_spat_M ==   True  ):
            $ 2474 "MoveJ" "noBreak"
            $ 2475 "Spatula_otw" "noBreak"
            movej(get_inverse_kin(Spatula_otw_p, qnear=Spatula_otw_q), a=1.3962634015954636, v=1.0471975511965976)
            $ 2476 "spat_L_up" "noBreak"
            movej(get_inverse_kin(spat_L_up_p, qnear=spat_L_up_q), a=1.3962634015954636, v=1.0471975511965976)
            $ 2477 "MoveL" "noBreak"
            $ 2478 "spat_L_side" "noBreak"
            movel(spat_L_side_p, a=1.2, v=0.25)
            $ 2479 "spat_L_lift" "noBreak"
            movel(spat_L_lift_p, a=1.2, v=0.25)
            $ 2480 "spat_L_pick" "noBreak"
            movel(spat_L_pick_p, a=1.2, v=0.25)
            # begin: URCap Program Node
            #   Source: Robotiq_Grippers, 1.8.4.4844, Robotiq Inc.
            #   Type: Gripper
            $ 2481 "Gripper Open (1)" "noBreak"
            if not(gripper_connected[0]):
              popup("Gripper 1 must be connected to run this program.", "No connection", False, True, True)
            end
            if not(rq_is_gripper_activated("1")):
              popup("Gripper 1 is not activated. Go to Installation tab > Gripper to activate it and run the program again.", "Not activated", False, True, True)
            end
            rq_set_pos_spd_for(0, 255, 77, "1")
            rq_wait_pos_spe_for_request(0, 255, 77, "1")
            rq_go_to("1")
            rq_wait("1")
            # end: URCap Program Node
            $ 2482 "spat_M_pick" "noBreak"
            movel(spat_M_pick_p, a=1.2, v=0.25)
            # begin: URCap Program Node
            #   Source: Robotiq_Grippers, 1.8.4.4844, Robotiq Inc.
            #   Type: Gripper
            $ 2483 "Gripper Close (1)" "noBreak"
            if not(gripper_connected[0]):
              popup("Gripper 1 must be connected to run this program.", "No connection", False, True, True)
            end
            if not(rq_is_gripper_activated("1")):
              popup("Gripper 1 is not activated. Go to Installation tab > Gripper to activate it and run the program again.", "Not activated", False, True, True)
            end
            rq_set_pos_spd_for(255, 0, 77, "1")
            rq_wait_pos_spe_for_request(255, 0, 77, "1")
            rq_go_to("1")
            rq_wait("1")
            # end: URCap Program Node
            $ 2484 "spat_M_up" "noBreak"
            movel(spat_M_up_p, a=1.2, v=0.25)
            $ 2485 "Spatula_otw" "noBreak"
            movel(Spatula_otw_p, a=1.2, v=0.25)
            $ 2486 "switch_spat_M≔ False " "noBreak"
            global switch_spat_M=  False
          else:
            $ 2487 "ElseIf spatula ≟ 'spatula_S' and switch_spat_S ≟ True " "noBreak"
            if (spatula  ==  "spatula_S" and switch_spat_S  ==   True  ):
              $ 2488 "MoveL" "noBreak"
              $ 2489 "Spatula_otw" "noBreak"
              movel(Spatula_otw_p, a=1.2, v=0.25)
              $ 2490 "spat_M_up" "noBreak"
              movel(spat_M_up_p, a=1.2, v=0.25)
              $ 2491 "spat_M_pick" "noBreak"
              movel(spat_M_pick_p, a=1.2, v=0.25)
              # begin: URCap Program Node
              #   Source: Robotiq_Grippers, 1.8.4.4844, Robotiq Inc.
              #   Type: Gripper
              $ 2492 "Gripper Open (1)" "noBreak"
              if not(gripper_connected[0]):
                popup("Gripper 1 must be connected to run this program.", "No connection", False, True, True)
              end
              if not(rq_is_gripper_activated("1")):
                popup("Gripper 1 is not activated. Go to Installation tab > Gripper to activate it and run the program again.", "Not activated", False, True, True)
              end
              rq_set_pos_spd_for(0, 255, 77, "1")
              rq_wait_pos_spe_for_request(0, 255, 77, "1")
              rq_go_to("1")
              rq_wait("1")
              # end: URCap Program Node
              $ 2493 "spat_S_pick" "noBreak"
              movel(spat_S_pick_p, a=1.2, v=0.25)
              # begin: URCap Program Node
              #   Source: Robotiq_Grippers, 1.8.4.4844, Robotiq Inc.
              #   Type: Gripper
              $ 2494 "Gripper Close (1)" "noBreak"
              if not(gripper_connected[0]):
                popup("Gripper 1 must be connected to run this program.", "No connection", False, True, True)
              end
              if not(rq_is_gripper_activated("1")):
                popup("Gripper 1 is not activated. Go to Installation tab > Gripper to activate it and run the program again.", "Not activated", False, True, True)
              end
              rq_set_pos_spd_for(255, 0, 77, "1")
              rq_wait_pos_spe_for_request(255, 0, 77, "1")
              rq_go_to("1")
              rq_wait("1")
              # end: URCap Program Node
              $ 2495 "spat_S_up" "noBreak"
              movel(spat_S_up_p, a=1.2, v=0.25)
              $ 2496 "Spatula_otw" "noBreak"
              movel(Spatula_otw_p, a=1.2, v=0.25)
              $ 2497 "switch_spat_S≔ False " "noBreak"
              global switch_spat_S=  False
            end
          end
          $ 2498 "auto_tilt_and_scoop(W_now, Target_weight, Weight_value)" "noBreak"
          auto_tilt_and_scoop(W_now, Target_weight, Weight_value)
          $ 2499 "Wait: 0.5" "noBreak"
          sleep(0.5)
        end
        # begin: URCap Program Node
        #   Source: SensoPart VISOR Robotic, 2.0.0, SensoPart Industriesensorik GmbH
        #   Type: Exit Pose
        $ 2501 "Exit Pose" "noBreak"
        movel(pose_trans(easyPickPose,p[0.0000,0.0000,-0.0000,0.0000,0.0000,0.0000]),a=0.5000,v=0.2500,t=0.000000,r=0.000000)
        # end: URCap Program Node
        easyPickObjTaken = True
      end
      # end: URCap Program Node
      # begin: URCap Program Node
      #   Source: SensoPart VISOR Robotic, 2.0.0, SensoPart Industriesensorik GmbH
      #   Type: No Object Detected
      $ 2502 "No Object Detected" "noBreak"
      if (visor_partsFound(easyPickVisorId) < 1):
        $ 2503 "Popup: No weigh scale detected" "noBreak"
        popup("No weigh scale detected", "Message", False, False, blocking=True)
        else:
      end
      # end: URCap Program Node
    end
    easyPickCount_4 = easyPickCount_4 + 1
    visor_easyPickUpdate(easyPickVisorId, "counter", easyPickCount_4)
    visor_easyPickSetIdent("7aa8bf", easyPickVisorId)
    # end: URCap Program Node
  end
  visorFuncEasyPick_221058()
  # end: URCap Program Node
  elif (42 == switch_1):
    $ 2566 "Case 42"
    $ 2567 "Powder dosing"
    $ 2568 "zero_scale()"
    zero_scale()
    $ 2569 "Task≔'Dosing'"
    global Task="Dosing"
    $ 2570 "scooping_init()"
    scooping_init()
    # begin: URCap Program Node
    #   Source: SensoPart VISOR Robotic, 2.0.0, SensoPart Industriesensorik GmbH
    #   Type: VISOR Robotic App
    $ 2571 "VISOR Easy Pick"
    def visorFuncEasyPick_68fcc5():
      # begin: URCap Program Node
      #   Source: SensoPart VISOR Robotic, 2.0.0, SensoPart Industriesensorik GmbH
      #   Type: Easy Pick Setup
      $ 2572 "# 1 Setup" "noBreak"
      local easyPickVisorId = 1
      local easyPickArmMounted = True
      local easyPickSetJob = True
      local easyPickJobName = "Weigh_target"
      local easyPickAtImgAcq = False
      local easyPickImgAcqPose = FRM_Weigh_scale
      # end: URCap Program Node
      # begin: URCap Program Node
      #   Source: SensoPart VISOR Robotic, 2.0.0, SensoPart Industriesensorik GmbH
      #   Type: Process
      $ 2573 "Process" "noBreak"
      local easyPickObjTaken = False
      local easyPickTrigger = False
      local easyPickPoseIdx = 0
      local easyPickPose = p[0,0,0,0,0,0]
      def easyPickFuncTrigger(visorId, setJob, jobName, arm):
      if (setJob):
        visor_changeJob(visorId, jobName, 6000)
      end
      if (arm):
        visor_trigger(visorId, 6000, "arm")
      else:
        visor_trigger(visorId, 6000)
      end
      global easyPickParts_4=visor_partsFound(visorId)
      visor_easyPickUpdate(visorId, "parts", visor_partsFound(visorId))
      return visor_getPose3d(visorId, 0)
    end
    while (not easyPickObjTaken):
      easyPickTrigger = (easyPickCount_4 >= visor_partsFound(easyPickVisorId)) or (easyPickCount_4 > 9) or (not visor_easyPickCheckIdent("14a4aa", easyPickVisorId))
      if (easyPickTrigger):
        easyPickCount_4 = 0
      end
      easyPickPoseIdx = easyPickCount_4
      easyPickPose = visor_getPose3d(easyPickVisorId, easyPickPoseIdx)
      visor_easyPickUpdate(easyPickVisorId, "counter", easyPickPoseIdx)
      # begin: URCap Program Node
      #   Source: SensoPart VISOR Robotic, 2.0.0, SensoPart Industriesensorik GmbH
      #   Type: Image Acquisition Pose
      $ 2574 "Image Acquisition Pose" "noBreak"
      if (easyPickTrigger):
        if (not easyPickAtImgAcq):
          movej(pose_trans(easyPickImgAcqPose,p[0.0000,0.0000,-0.0000,0.0000,0.0000,0.0000]),a=1.3963,v=1.0472,t=0.000000,r=0.000000)
          easyPickAtImgAcq = True
        end
        easyPickPose = easyPickFuncTrigger(easyPickVisorId, easyPickSetJob, easyPickJobName, easyPickArmMounted)
      end
      # end: URCap Program Node
      # begin: URCap Program Node
      #   Source: SensoPart VISOR Robotic, 2.0.0, SensoPart Industriesensorik GmbH
      #   Type: Object Detected
      $ 2575 "Object Detected" "noBreak"
      if (visor_partsFound(easyPickVisorId) > 0):
        $ 2576 "Open Gripper" "noBreak"
        $ 2577 "tare_scale()" "noBreak"
        tare_scale()
        $ 2578 "Wait: 0.2" "noBreak"
        sleep(0.2)
        $ 2579 "Weight_value≔get_weight()" "noBreak"
        global Weight_value=get_weight()
        $ 2580 "Wait: 0.2" "noBreak"
        sleep(0.2)
        $ 2581 "diff≔Target_weight-Weight_value" "noBreak"
        global diff=Target_weight-Weight_value
        $ 2582 "compute_level_percent(W_now, Weight_value)" "noBreak"
        compute_level_percent(W_now, Weight_value)
        $ 2583 "spatula = select_spatula(Pow_name, level, diff)" "noBreak"
        spatula = select_spatula(Pow_name, level, diff)
        $ 2584 "If spatula ≟ 'spatula_L'" "noBreak"
        if (spatula  ==  "spatula_L"):
          $ 2585 "MoveJ" "noBreak"
          $ 2586 "Spatula_otw" "noBreak"
          movej(get_inverse_kin(Spatula_otw_p, qnear=Spatula_otw_q), a=1.3962634015954636, v=1.0471975511965976)
          $ 2587 "pick_spat_L_abv" "noBreak"
          movej(get_inverse_kin(pick_spat_L_abv_p, qnear=pick_spat_L_abv_q), a=1.3962634015954636, v=1.0471975511965976)
          $ 2588 "MoveL" "noBreak"
          $ 2589 "spat_L_pick" "noBreak"
          movel(spat_L_pick_p, a=1.2, v=0.25)
          # begin: URCap Program Node
          #   Source: Robotiq_Grippers, 1.8.4.4844, Robotiq Inc.
          #   Type: Gripper
          $ 2590 "Gripper Close (1)" "noBreak"
          if not(gripper_connected[0]):
            popup("Gripper 1 must be connected to run this program.", "No connection", False, True, True)
          end
          if not(rq_is_gripper_activated("1")):
            popup("Gripper 1 is not activated. Go to Installation tab > Gripper to activate it and run the program again.", "Not activated", False, True, True)
          end
          rq_set_pos_spd_for(255, 0, 77, "1")
          rq_wait_pos_spe_for_request(255, 0, 77, "1")
          rq_go_to("1")
          rq_wait("1")
          # end: URCap Program Node
          $ 2591 "spat_L_lift" "noBreak"
          movel(spat_L_lift_p, a=1.2, v=0.25)
          $ 2592 "spat_L_side" "noBreak"
          movel(spat_L_side_p, a=1.2, v=0.25)
          $ 2593 "spat_L_up" "noBreak"
          movel(spat_L_up_p, a=1.2, v=0.25)
          $ 2594 "MoveJ" "noBreak"
          $ 2595 "Spatula_otw" "noBreak"
          movej(get_inverse_kin(Spatula_otw_p, qnear=Spatula_otw_q), a=1.3962634015954636, v=1.0471975511965976)
        else:
          $ 2596 "ElseIf spatula ≟'spatula_M'" "noBreak"
          if (spatula  == "spatula_M"):
            $ 2597 "MoveJ" "noBreak"
            $ 2598 "Spatula_otw" "noBreak"
            movej(get_inverse_kin(Spatula_otw_p, qnear=Spatula_otw_q), a=1.3962634015954636, v=1.0471975511965976)
            $ 2599 "spat_M_up" "noBreak"
            movej(get_inverse_kin(spat_M_up_p, qnear=spat_M_up_q), a=1.3962634015954636, v=1.0471975511965976)
            $ 2600 "MoveL" "noBreak"
            $ 2601 "spat_M_pick" "noBreak"
            movel(spat_M_pick_p, a=1.2, v=0.25)
            # begin: URCap Program Node
            #   Source: Robotiq_Grippers, 1.8.4.4844, Robotiq Inc.
            #   Type: Gripper
            $ 2602 "Gripper Close (1)" "noBreak"
            if not(gripper_connected[0]):
              popup("Gripper 1 must be connected to run this program.", "No connection", False, True, True)
            end
            if not(rq_is_gripper_activated("1")):
              popup("Gripper 1 is not activated. Go to Installation tab > Gripper to activate it and run the program again.", "Not activated", False, True, True)
            end
            rq_set_pos_spd_for(255, 0, 77, "1")
            rq_wait_pos_spe_for_request(255, 0, 77, "1")
            rq_go_to("1")
            rq_wait("1")
            # end: URCap Program Node
            $ 2603 "spat_M_up" "noBreak"
            movel(spat_M_up_p, a=1.2, v=0.25)
            $ 2604 "Spatula_otw" "noBreak"
            movel(Spatula_otw_p, a=1.2, v=0.25)
            $ 2605 "switch_spat_M≔ False " "noBreak"
            global switch_spat_M=  False
          else:
            $ 2606 "ElseIf spatula≟'spatula_S'" "noBreak"
            if (spatula == "spatula_S"):
              $ 2607 "MoveJ" "noBreak"
              $ 2608 "Spatula_otw" "noBreak"
              movej(get_inverse_kin(Spatula_otw_p, qnear=Spatula_otw_q), a=1.3962634015954636, v=1.0471975511965976)
              $ 2609 "spat_M_up" "noBreak"
              movej(get_inverse_kin(spat_M_up_p, qnear=spat_M_up_q), a=1.3962634015954636, v=1.0471975511965976)
              $ 2610 "MoveL" "noBreak"
              $ 2611 "spat_M_pick" "noBreak"
              movel(spat_M_pick_p, a=1.2, v=0.25)
              # begin: URCap Program Node
              #   Source: Robotiq_Grippers, 1.8.4.4844, Robotiq Inc.
              #   Type: Gripper
              $ 2612 "Gripper Close (1)" "noBreak"
              if not(gripper_connected[0]):
                popup("Gripper 1 must be connected to run this program.", "No connection", False, True, True)
              end
              if not(rq_is_gripper_activated("1")):
                popup("Gripper 1 is not activated. Go to Installation tab > Gripper to activate it and run the program again.", "Not activated", False, True, True)
              end
              rq_set_pos_spd_for(255, 0, 77, "1")
              rq_wait_pos_spe_for_request(255, 0, 77, "1")
              rq_go_to("1")
              rq_wait("1")
              # end: URCap Program Node
              $ 2613 "spat_M_up" "noBreak"
              movel(spat_M_up_p, a=1.2, v=0.25)
              $ 2614 "Spatula_otw" "noBreak"
              movel(Spatula_otw_p, a=1.2, v=0.25)
              $ 2615 "switch_spat_M≔ False " "noBreak"
              global switch_spat_M=  False
            end
          end
        end
        $ 2616 "Weight_value≔get_weight()" "noBreak"
        global Weight_value=get_weight()
        $ 2617 "auto_tilt_and_scoop(W_now, Target_weight, Weight_value)" "noBreak"
        auto_tilt_and_scoop(W_now, Target_weight, Weight_value)
        # begin: URCap Program Node
        #   Source: SensoPart VISOR Robotic, 2.0.0, SensoPart Industriesensorik GmbH
        #   Type: Approach Pose
        $ 2618 "Approach Pose" "noBreak"
        movej(pose_trans(easyPickPose,p[0.0000,0.0000,0.0500,0.0000,0.0000,0.0000]),a=0.2618,v=0.1745,t=0.000000,r=0.000000)
        # end: URCap Program Node
        # begin: URCap Program Node
        #   Source: SensoPart VISOR Robotic, 2.0.0, SensoPart Industriesensorik GmbH
        #   Type: Target Pose
        $ 2619 "Target Pose" "noBreak"
        movel(pose_trans(easyPickPose,p[0.0000,0.0000,-0.0000,0.0000,0.0000,0.0000]),a=0.0500,v=0.0200,t=0.000000,r=0.000000)
        # end: URCap Program Node
        $ 2620 "Close Gripper" "noBreak"
        $ 2621 "dispense_pos≔get_actual_tcp_pose()" "noBreak"
        global dispense_pos= get_actual_tcp_pose ()
        $ 2622 "Loop Weight_value≤Target_weight" "noBreak"
        thread Thread_while_2622():
          while (True):
            $ 2623 "MoveL" "noBreak"
            $ 2624 "dispense_pos" "noBreak"
            movel(dispense_pos, a=0.2, v=0.1)
            $ 2625 "log_weight()" "noBreak"
            log_weight()
            $ 2626 "Wait: 0.5" "noBreak"
            sleep(0.5)
            $ 2627 "If level≥90.0" "noBreak"
            if (level >= 90.0):
              $ 2628 "Rotate()" "noBreak"
              Rotate()
            end
            $ 2629 "If level≤70" "noBreak"
            if (level <= 70):
              $ 2630 "tilt_to_home()" "noBreak"
              tilt_to_home()
            end
            $ 2631 "Wait: 0.5" "noBreak"
            sleep(0.5)
            $ 2632 "Start_thread≔ True " "noBreak"
            global Start_thread=  True
            $ 2633 "vib_mot_thread≔ True " "noBreak"
            global vib_mot_thread=  True
            $ 2635 "Wait: 0.5" "noBreak"
            sleep(0.5)
            $ 2641 "If spatula ≟ 'spatula_L'  and diff ≥3.5" "noBreak"
            if (spatula  ==  "spatula_L"   and  diff  >= 3.5):
              $ 2642 "tilt_pose≔pose_trans(get_actual_tcp_pose(), p[0, 0, 0, 0, 0, 2.0])" "noBreak"
              global tilt_pose=pose_trans(get_actual_tcp_pose(), p[0, 0, 0, 0, 0, 2.0])
              $ 2643 "movel(tilt_pose, a=0.1, v=0.1, r=0.00001)" "noBreak"
              movel(tilt_pose, a=0.1, v=0.1, r=0.00001)
            end
            $ 2655 "If spatula ≟ 'spatula_M'  and diff ≥1.0" "noBreak"
            if (spatula  ==  "spatula_M"   and  diff  >= 1.0):
              $ 2656 "tilt_pose≔pose_trans(get_actual_tcp_pose(), p[0, 0, 0, 0, 0, 2.0])" "noBreak"
              global tilt_pose=pose_trans(get_actual_tcp_pose(), p[0, 0, 0, 0, 0, 2.0])
              $ 2657 "movel(tilt_pose, a=0.1, v=0.1, r=0.00001)" "noBreak"
              movel(tilt_pose, a=0.1, v=0.1, r=0.00001)
            else:
              $ 2658 "ElseIf diff≤1.0" "noBreak"
              if (diff <= 1.0):
                $ 2659 "Loop Weight_value≤Target_weight and tilt_angle≥(-1.999) and tilt_angle≤0.5" "noBreak"
                while (Weight_value <= Target_weight  and  tilt_angle >= (-1.999)  and  tilt_angle <= 0.5):
                  $ 2660 "current_error≔Target_weight-Weight_value" "noBreak"
                  global current_error=Target_weight-Weight_value
                  $ 2661 "Integral_error≔Integral_error+current_error*dt" "noBreak"
                  global Integral_error=Integral_error+current_error*dt
                  $ 2662 "derivative≔(current_error-previous_error)/dt" "noBreak"
                  global derivative=(current_error-previous_error)/dt
                  $ 2663 "tilt_increment≔(kp*current_error)+(ki*Integral_error)+(kd*derivative)" "noBreak"
                  global tilt_increment=(kp*current_error)+(ki*Integral_error)+(kd*derivative)
                  $ 2664 "current_pose≔get_actual_tcp_pose()" "noBreak"
                  global current_pose= get_actual_tcp_pose ()
                  $ 2665 "tilt_angle≔current_pose[5]" "noBreak"
                  global tilt_angle=current_pose[5]
                  $ 2666 "tilt_pose≔pose_trans(current_pose, p[0, 0, 0, 0, 0, tilt_increment])" "noBreak"
                  global tilt_pose=pose_trans(current_pose, p[0, 0, 0, 0, 0, tilt_increment])
                  $ 2667 "movel(tilt_pose, a=0.1, v=0.1, r=0.00001)" "noBreak"
                  movel(tilt_pose, a=0.1, v=0.1, r=0.00001)
                  $ 2668 "previous_error≔current_error" "noBreak"
                  global previous_error=current_error
                end
              end
            end
            $ 2669 "Start_thread≔ False " "noBreak"
            global Start_thread=  False
            $ 2671 "Weight_value≔get_weight()" "noBreak"
            global Weight_value=get_weight()
            $ 2673 "Wait: 0.5" "noBreak"
            sleep(0.5)
            $ 2674 "vib_mot_thread≔ False " "noBreak"
            global vib_mot_thread=  False
            $ 2675 "MoveL" "noBreak"
            $ 2676 "dispense_pos" "noBreak"
            movel(dispense_pos, a=0.5, v=0.25)
            $ 2677 "Integral_error≔0" "noBreak"
            global Integral_error=0
            $ 2678 "current_error≔0" "noBreak"
            global current_error=0
            $ 2679 "previous_error≔0" "noBreak"
            global previous_error=0
            $ 2680 "Set AO[0]=0.0" "noBreak"
            set_standard_analog_out(0, 0.0)
            $ 2681 "select_spatula(Pow_name, level, diff)" "noBreak"
            select_spatula(Pow_name, level, diff)
            $ 2682 "If spatula ≟ 'spatula_M'  and switch_spat_M≟ True " "noBreak"
            if (spatula  ==  "spatula_M"   and  switch_spat_M ==   True  ):
              $ 2683 "MoveJ" "noBreak"
              $ 2684 "Spatula_otw" "noBreak"
              movej(get_inverse_kin(Spatula_otw_p, qnear=Spatula_otw_q), a=1.3962634015954636, v=1.0471975511965976)
              $ 2685 "spat_L_up" "noBreak"
              movej(get_inverse_kin(spat_L_up_p, qnear=spat_L_up_q), a=1.3962634015954636, v=1.0471975511965976)
              $ 2686 "MoveL" "noBreak"
              $ 2687 "spat_L_side" "noBreak"
              movel(spat_L_side_p, a=1.2, v=0.25)
              $ 2688 "spat_L_lift" "noBreak"
              movel(spat_L_lift_p, a=1.2, v=0.25)
              $ 2689 "spat_L_pick" "noBreak"
              movel(spat_L_pick_p, a=1.2, v=0.25)
              # begin: URCap Program Node
              #   Source: Robotiq_Grippers, 1.8.4.4844, Robotiq Inc.
              #   Type: Gripper
              $ 2690 "Gripper Open (1)" "noBreak"
              if not(gripper_connected[0]):
                popup("Gripper 1 must be connected to run this program.", "No connection", False, True, True)
              end
              if not(rq_is_gripper_activated("1")):
                popup("Gripper 1 is not activated. Go to Installation tab > Gripper to activate it and run the program again.", "Not activated", False, True, True)
              end
              rq_set_pos_spd_for(0, 255, 77, "1")
              rq_wait_pos_spe_for_request(0, 255, 77, "1")
              rq_go_to("1")
              rq_wait("1")
              # end: URCap Program Node
              $ 2691 "spat_M_pick" "noBreak"
              movel(spat_M_pick_p, a=1.2, v=0.25)
              # begin: URCap Program Node
              #   Source: Robotiq_Grippers, 1.8.4.4844, Robotiq Inc.
              #   Type: Gripper
              $ 2692 "Gripper Close (1)" "noBreak"
              if not(gripper_connected[0]):
                popup("Gripper 1 must be connected to run this program.", "No connection", False, True, True)
              end
              if not(rq_is_gripper_activated("1")):
                popup("Gripper 1 is not activated. Go to Installation tab > Gripper to activate it and run the program again.", "Not activated", False, True, True)
              end
              rq_set_pos_spd_for(255, 0, 77, "1")
              rq_wait_pos_spe_for_request(255, 0, 77, "1")
              rq_go_to("1")
              rq_wait("1")
              # end: URCap Program Node
              $ 2693 "spat_M_up" "noBreak"
              movel(spat_M_up_p, a=1.2, v=0.25)
              $ 2694 "Spatula_otw" "noBreak"
              movel(Spatula_otw_p, a=1.2, v=0.25)
              $ 2695 "switch_spat_M≔ False " "noBreak"
              global switch_spat_M=  False
            else:
              $ 2696 "ElseIf spatula ≟ 'spatula_S' and switch_spat_S ≟ True " "noBreak"
              if (spatula  ==  "spatula_S" and switch_spat_S  ==   True  ):
                $ 2697 "MoveL" "noBreak"
                $ 2698 "Spatula_otw" "noBreak"
                movel(Spatula_otw_p, a=1.2, v=0.25)
                $ 2699 "spat_M_up" "noBreak"
                movel(spat_M_up_p, a=1.2, v=0.25)
                $ 2700 "spat_M_pick" "noBreak"
                movel(spat_M_pick_p, a=1.2, v=0.25)
                # begin: URCap Program Node
                #   Source: Robotiq_Grippers, 1.8.4.4844, Robotiq Inc.
                #   Type: Gripper
                $ 2701 "Gripper Open (1)" "noBreak"
                if not(gripper_connected[0]):
                  popup("Gripper 1 must be connected to run this program.", "No connection", False, True, True)
                end
                if not(rq_is_gripper_activated("1")):
                  popup("Gripper 1 is not activated. Go to Installation tab > Gripper to activate it and run the program again.", "Not activated", False, True, True)
                end
                rq_set_pos_spd_for(0, 255, 77, "1")
                rq_wait_pos_spe_for_request(0, 255, 77, "1")
                rq_go_to("1")
                rq_wait("1")
                # end: URCap Program Node
                $ 2702 "spat_S_pick" "noBreak"
                movel(spat_S_pick_p, a=1.2, v=0.25)
                # begin: URCap Program Node
                #   Source: Robotiq_Grippers, 1.8.4.4844, Robotiq Inc.
                #   Type: Gripper
                $ 2703 "Gripper Close (1)" "noBreak"
                if not(gripper_connected[0]):
                  popup("Gripper 1 must be connected to run this program.", "No connection", False, True, True)
                end
                if not(rq_is_gripper_activated("1")):
                  popup("Gripper 1 is not activated. Go to Installation tab > Gripper to activate it and run the program again.", "Not activated", False, True, True)
                end
                rq_set_pos_spd_for(255, 0, 77, "1")
                rq_wait_pos_spe_for_request(255, 0, 77, "1")
                rq_go_to("1")
                rq_wait("1")
                # end: URCap Program Node
                $ 2704 "spat_S_up" "noBreak"
                movel(spat_S_up_p, a=1.2, v=0.25)
                $ 2705 "Spatula_otw" "noBreak"
                movel(Spatula_otw_p, a=1.2, v=0.25)
                $ 2706 "switch_spat_S≔ False " "noBreak"
                global switch_spat_S=  False
              end
            end
            $ 2707 "auto_tilt_and_scoop(W_now, Target_weight, Weight_value)" "noBreak"
            auto_tilt_and_scoop(W_now, Target_weight, Weight_value)
            $ 2708 "Wait: 0.5" "noBreak"
            sleep(0.5)
          end
        end
        if (Weight_value <= Target_weight):
          global thread_handler_2622=run Thread_while_2622()
          while (Weight_value <= Target_weight):
            sync()
          end
          kill thread_handler_2622
        end
        $ 2709 "Start_thread≔ False " "noBreak"
        global Start_thread=  False
        $ 2710 "Wait: 0.5" "noBreak"
        sleep(0.5)
        $ 2711 "vib_mot_thread≔ False " "noBreak"
        global vib_mot_thread=  False
        # begin: URCap Program Node
        #   Source: SensoPart VISOR Robotic, 2.0.0, SensoPart Industriesensorik GmbH
        #   Type: Exit Pose
        $ 2713 "Exit Pose" "noBreak"
        movel(pose_trans(easyPickPose,p[0.0000,0.0000,-0.0000,0.0000,0.0000,0.0000]),a=0.5000,v=0.2500,t=0.000000,r=0.000000)
        # end: URCap Program Node
        easyPickObjTaken = True
      end
      # end: URCap Program Node
      # begin: URCap Program Node
      #   Source: SensoPart VISOR Robotic, 2.0.0, SensoPart Industriesensorik GmbH
      #   Type: No Object Detected
      $ 2714 "No Object Detected" "noBreak"
      if (visor_partsFound(easyPickVisorId) < 1):
        $ 2715 "Popup: No weigh scale detected" "noBreak"
        popup("No weigh scale detected", "Message", False, False, blocking=True)
        else:
      end
      # end: URCap Program Node
    end
    easyPickCount_4 = easyPickCount_4 + 1
    visor_easyPickUpdate(easyPickVisorId, "counter", easyPickCount_4)
    visor_easyPickSetIdent("14a4aa", easyPickVisorId)
    # end: URCap Program Node
  end
  visorFuncEasyPick_68fcc5()
  # end: URCap Program Node
  $ 2716 "MoveJ"
  $ 2717 "dispense_pos" "breakAfter"
  movej(dispense_pos, a=0.5235987755982988, v=0.4363323129985824)
  $ 2718 "after_scoop()"
  after_scoop()
  end
  $ 2781 "'=========='"
  # '=========='
  $ 2782 "PostSettings"
  $ 2783 "'ADD ADDITIONAL CHECKS'"
  # 'ADD ADDITIONAL CHECKS'
  end
  $ 2 "BeforeStart"
  $ 3 "Scripts"
  $ 4 "Script: 001 SCRIPT Errors and Warnings Deifnes V0.2.script"

  #*****************************************************
  # customer          :   UK Essen
  # project name      :   P1132
  #****************************************************
  # controller        :
  # software          :
  #****************************************************
  # author            :   E.Petrichenko
  # Copyright (c)     :   United Robotics Group Health and Food GmbH
  #                       An der Riede 2
  #                       28816 Stuhr
  #                       Germany
  #****************************************************
  # description       :   centrifuge actions for the application
  # version:      	:   0.1
  # created           :   22.08.2024
  # updated           :
  #****************************************************
  # modifications     :
  #
  # date              :
  # name              :
  # reason            :
  #****************************************************


  #################################### VARIABLES DEFINITIONS ###################################

  ERROR_POSE_NOT_REACHABLE = 1002
  ERROR_ROBOT_ARM_NOT_IN_HOME_POSE = 1006
  ERROR_NO_OBJECT_TO_PICK = 1010
  ERROR_NOT_DOCKED = 2003
  ERROR_NOT_REACHABLE_TARGET = 2007
  ERROR_CHARGING_NOT_STARTED = 2008
  ERROR_AMR_WRONG_MODE = 2009
  ERROR_UNKNOWN_POSE = 2010
  ERROR_NO_LANDMARK = 3002
  ERROR_WRONG_ORDER = 4002
  ERROR_CENTRIFUGE_CONNECTION = 5001
  ERROR_CENTRIFUGE_POWER = 5002
  ERROR_CENTRIFUGE = 5003
  ERROR_CENTRIFUGE_LID = 5004
  ERROR_CANNOT_OPEN_HATCH = 5006
  ERROR_CANNOT_CLOSE_HATCH = 5008
  ERROR_CANNOT_ROTATE = 5010
  ERROR_CANNOT_START = 5011
  ERROR_WRONG_KEY_POSE = 5012
  ERROR_MISSIING_CENTRACK = 5013

  WARNING_POSE_NOT_REACHABLE = 1002
  WARNING_BATTERY_LEVEL = 2002
  WARNING_NOT_REACHABLE_TARGET = 2007


  ERROR = struct(
      FLAG = False,
      ID = 0,
      MSG = "")

  WARNING = struct(
      FLAG = False,
      ID = 0,
      MSG = "")


  #################################### FUNCTIONS ###################################

  def set_error(error_id):
      ERROR.ID = error_id
      if (ERROR.ID == 0):
          ERROR.FLAG = False
          ERROR.MSG = ""
      else:
          ERROR.FLAG = True
          if(ERROR.ID == ERROR_POSE_NOT_REACHABLE):
              ERROR.MSG = "Pose is not reachable"
          elif(ERROR.ID == ERROR_NO_OBJECT_TO_PICK):
              ERROR.MSG = "No object to pick"
          elif(ERROR.ID == ERROR_NO_LANDMARK):
              ERROR.MSG = "No landmark detected"
          elif(ERROR.ID == ERROR_ROBOT_ARM_NOT_IN_HOME_POSE):
              ERROR.MSG = "Robot arm cannot go to home pose"
          elif(ERROR.ID == ERROR_AMR_WRONG_MODE):
              ERROR.MSG = "AMR is in the wrong mode"
          elif(ERROR.ID == ERROR_NOT_DOCKED):
              ERROR.MSG = "Could not dock to the charger"
          elif(ERROR.ID == ERROR_NOT_REACHABLE_TARGET):
              ERROR.MSG = "Could not reach the target"
          elif(ERROR.ID == ERROR_CHARGING_NOT_STARTED):
              ERROR.MSG = "Could not start charging"
          elif(ERROR.ID == ERROR_UNKNOWN_POSE):
              ERROR.MSG = "Unknown navigation target"
          elif(ERROR.ID == ERROR_CANNOT_OPEN_HATCH):
              ERROR.MSG = "Centrifuge Cannot open the hatch"
          elif(ERROR.ID == ERROR_CENTRIFUGE_CONNECTION):
              ERROR.MSG = "Cannot reach centrifuge"
          elif (ERROR.ID == ERROR_CANNOT_CLOSE_HATCH):
              ERROR.MSG = "Centrifuge Cannot close the hatch"
          elif (ERROR.ID == ERROR_CANNOT_START):
              ERROR.MSG = "Centrifuge Cannot start"
          elif (ERROR.ID == ERROR_CANNOT_ROTATE):
              ERROR.MSG = "Centrifuge Cannot rotate the rotor"
          elif (ERROR.ID == ERROR_WRONG_ORDER):
              ERROR.MSG = "Wrong parameter was recieved"
          elif (ERROR.ID == ERROR_CENTRIFUGE):
              ERROR.MSG = "Centrifuge is in Error"
          elif (ERROR.ID == ERROR_WRONG_KEY_POSE):
              ERROR.MSG = "Key is in the wrong position"
          elif(ERROR.ID == ERROR_MISSIING_CENTRACK):
              ERROR.MSG = "Missing rack for centrifuge set"
          elif(ERROR.ID == ERROR_CENTRIFUGE_POWER):
              ERROR.MSG = "Centrifuge is turned off"
          elif(ERROR.ID == ERROR_CENTRIFUGE_LID):
              ERROR.MSG = "Lid of the centrifuge is opened"
          else:
              ERROR.MSG = "Unknown code"
          end
          textmsg("ERROR:",ERROR)
      end
  end

  def set_warning(warning_id):
      WARNING.ID = warning_id
      if (WARNING.ID == 0):
          WARNING.FLAG = False
          WARNING.MSG = ""
      else:
          WARNING.FLAG = True
          if(WARNING.ID == WARNING_POSE_NOT_REACHABLE):
              WARNING.MSG = "Pose is not reachable"
          elif(WARNING.ID == WARNING_BATTERY_LEVEL):
              WARNING.MSG = "Batery level dropped to a certain level"
          elif(WARNING.ID == WARNING_NOT_REACHABLE_TARGET):
              WARNING.MSG = "Not reachable location of AMR"
          else:
              WARNING.MSG = "Unknown code"
          end
          textmsg("WARNING:",WARNING)
      end
  end


  def reset_error():
    ERROR.ID = 0
    ERROR.FLAG = False
    ERROR.MSG = ""
  end


  def reset_warning():
      WARNING.ID = 0
      WARNING.FLAG = False
      WARNING.MSG = ""
    end
  $ 5 "Script: SCRIPT uGO V7.11.1.script"
  #*****************************************************
  # customer          :
  # project name      :   Standard Application
  #****************************************************
  # controller        :
  # software          :
  #****************************************************
  # author            :   P. Koehnke
  # Copyright (c)     :   United Robotics Group
  #                       An der Riede 2
  #                       28816 Stuhr
  #                       Germany
  #****************************************************
  # description       :   interface for uGo
  # version:      	:   6.0
  # created           :   21.04.2022
  # updated           :
  #****************************************************
  # modifications     :   add new rpc-functions to interchange more data
  #
  # date              :   2024-02-29
  # name              :   P. Koehnke
  # reason            :   implemtentation of PackML behavoiur in uGO
  #****************************************************
  #****************************************************
  # modifications     :   add reflecting the UID of the uGO task back to uGO
  #
  # date              :   2024-07-02
  # name              :   P. Koehnke
  # reason            :   be sure to finish the right tasks
  #****************************************************

  # available rpc-functions:
  #.on('con_check', (err, _params, callback) => callback(err, this.con_check()))
  #.on('read_input', (err, params, callback) => callback(err, this.read_input(params[0], params[1])))
  #.on('write_output', (err, params, callback) => callback(err, this.write_output(params[0], params[1], params[2])))
  #.on('read_status', (err, params, callback) => callback(err, this.read_status(params[0])))
  #.on('write_status', (err, params, callback) => callback(err, this.write_status(params[0], params[1])))
  #.on('send_template', (err, params, callback) => callback(err, this.receive_state(params[0])))
  #.on('receive_event', (err, params, callback) => callback(err, this.send_event()))
  #.on('send_state', (err, params, callback) => callback(err, this.receive_state(params[0])))
  #.on('send_error', (err, params, callback) => callback(err, this.receive_error(params[0])))
  #.on('NotFound', (methodCalled, params) => LOG.warn('Method "', methodCalled, '" does not exist. ', { params }));

  # =======================================================================
  local IDX_CMD_STOP = 0
  local IDX_CMD_RESET = 1
  local IDX_CMD_START = 2
  local IDX_CMD_HOLD = 3
  local IDX_CMD_UNHOLD = 4
  local IDX_CMD_SUSPEND = 5
  local IDX_CMD_UNSUSPEND = 6
  local IDX_CMD_ABORT = 7
  local IDX_CMD_CLEAR = 8
  local IDX_FNC_FREEDRIVE = 9

  # uGo specific declarations
  global UGO_Request_ID = ""
  global UGO_UNIT_Task = ""
  global UGO_Task_ID = 0
  global UGO_Event = ""
  local UGO_Enable_Control = False
  local UGO = rpc_factory("xmlrpc", "http://192.168.12.120:8080")
  local UGO_Ctrl_Cmd = [False, False, False, False, False, False, False, False, False, False]

  local UGO_AMR_Pos = struct(position_identifier=0, x1=0, x2=0, y1=0, y2=0, theta1=0, theta2=0)
  local UGO_EOAT = struct(object_picked=False)

  def ugo_init(enable=True, rpc_address="http://192.168.12.120:8080"):
      # connection with uGo
      if enable:
          UGO = rpc_factory("xmlrpc", rpc_address)
          UGO_Enable_Control = True
      else:
          UGO_Enable_Control = False
      end
  end

  def ugo_event_controller():
      # interpret the given command and map it to the internal commands
      if UGO_Enable_Control:
          UGO_Event = UGO.receive_event()
      end

      UGO_Ctrl_Cmd[IDX_CMD_STOP] = (UGO_Event == "stop")
      UGO_Ctrl_Cmd[IDX_CMD_RESET] = (UGO_Event == "reset")
      UGO_Ctrl_Cmd[IDX_CMD_START] = (UGO_Event == "start")
      UGO_Ctrl_Cmd[IDX_CMD_HOLD] = (UGO_Event == "hold")
      UGO_Ctrl_Cmd[IDX_CMD_UNHOLD] = (UGO_Event == "un_hold")
      UGO_Ctrl_Cmd[IDX_CMD_SUSPEND] = (UGO_Event == "suspend")
      UGO_Ctrl_Cmd[IDX_CMD_UNSUSPEND] = (UGO_Event == "un_suspend")
      UGO_Ctrl_Cmd[IDX_CMD_ABORT] = (UGO_Event == "abort")
      UGO_Ctrl_Cmd[IDX_CMD_CLEAR] = (UGO_Event == "clear")
      UGO_Ctrl_Cmd[IDX_FNC_FREEDRIVE] = (UGO_Event == "freedrive")

      return UGO_Ctrl_Cmd
  end

  def ugo_translate_pml_state():
      # translate the current PML State to a string
      if (STATE == 1):
          return "STOPPING"
      elif (STATE == 2):
          return "STOPPED"
      elif (STATE == 3):
          return "RESETTING"
      elif (STATE == 4):
          return "IDLE"
      elif (STATE == 5):
          return "STARTING"
      elif (STATE == 6):
          return "EXECUTE"
      elif (STATE == 7):
          return "COMPLETING"
      elif (STATE == 8):
          return "COMPLETE"
      elif (STATE == 9):
          return "HOLDING"
      elif (STATE == 10):
          return "HELD"
      elif (STATE == 11):
          return "UNHOLDING"
      elif (STATE == 12):
          return "SUSPENDING"
      elif (STATE == 13):
          return "SUSPENDED"
      elif (STATE == 14):
          return "UNSUSPENDING"
      elif (STATE == 15):
          return "ABORTING"
      elif (STATE == 16):
          return "ABORTED"
      elif (STATE == 17):
          return "CLEARING"
      else:
          return "UNKNOWN"
      end
  end

  def ugo_update_outputs():
      #Update the outputs to uGo via xmplrpc service
      UGO.write_status("ROB_Skill", UGO_UNIT_Task)
      UGO.write_status("ROB_Battery", AMR_Battery)
      UGO.write_status("ROB_Gripper", OBJ_Picked)
      UGO.send_state(ugo_translate_pml_state(), UGO_UNIT_Task)
      UGO.send_error(ERROR.ID)
      #UGO.send_position(AMR_Position)
  end

  def ugo_get_task():
      # get the actual task to work on
      # added: reflecting the UID of the task back to uGO
      UGO_UNIT_Task = UGO.read_status("DSH_Workflow")
      if (UGO_UNIT_Task != ""):
          UGO_Request_ID = str_sub(UGO_UNIT_Task, 0, 39)
          UGO_Task_ID = to_num(str_sub(UGO_UNIT_Task, 40, 2))
          #ugo_tasks()
          return UGO_Task_ID
      else:
          return 0
      end
  end

  def ugo_pml_stopping():
      return True
  end

  def ugo_pml_resetting():
      ugo_get_task()
      if (UGO_UNIT_Task == ""):
          UGO_Request_ID = ""
          UGO_Task_ID = 0
          return True
      end
      return False
  end

  def ugo_pml_starting():
      #UGO_Task_Content = UGO.receive_task()
      return (UGO_UNIT_Task != "")
  end

  def ugo_pml_holding():
      return True
  end

  def ugo_pml_unholding():
      return True
  end

  def ugo_pml_suspending():
      return True
  end

  def ugo_pml_unsuspending():
      return True
  end

  def ugo_pml_completing():
      return True
  end

  def ugo_pml_aborting():
      return True
  end

  def ugo_pml_clearing():
      return True
  end

  # =======================================================================
  # end of uGO script
  # =======================================================================
  $ 7 "Script: SCRIPT PackML V1.2.1.script"
  # PackML

  IO_ADDRESS_CMD_STOP = 1
  IO_ADDRESS_CMD_RESET = 7
  IO_ADDRESS_CMD_START = 0

  EXT_ADDRESS_CMD_STOP = 0
  EXT_ADDRESS_CMD_RESET = 1
  EXT_ADDRESS_CMD_START = 2
  EXT_ADDRESS_CMD_HOLD = 3
  EXT_ADDRESS_CMD_UNHOLD = 4
  EXT_ADDRESS_CMD_SUSPEND = 5
  EXT_ADDRESS_CMD_UNSUSPEND = 6
  EXT_ADDRESS_CMD_ABORT = 7
  EXT_ADDRESS_CMD_CLEAR = 8
  EXT_ADDRESS_FNC_FREEDRIVE = 9

  global EXT_CtrlCmd = [False, False, False, False, False, False, False, False, False, False]

  EXT_Control_by = "uGO"

  global CMD_Abort = False
  global CMD_Clear = False
  global CMD_Stop = False
  global CMD_Reset = False
  global CMD_Start = False
  global CMD_Hold = False
  global CMD_Unhold = False
  global CMD_Suspend = False
  global CMD_Unsuspend = False
  global FNC_Freedrive = False

  CND_Suspend = False         # condition for suspend command
  CND_Unsuspend = False       # condition for unsuspend command

  thread Get_Pml_Command():
      while (True):
          if (EXT_Control_by == "uGO"):
              EXT_CtrlCmd = ugo_event_controller()
          elif (EXT_Control_by == "Leitsystem"):
              # EXT_CtrlCmd = Leitsystem
          end
          # ---------- Abort ---------- #
          if ((not STATE == 15) and (not STATE == 16) and EXT_CtrlCmd[EXT_ADDRESS_CMD_ABORT]):
              CMD_Abort = True
              CMD_Stop = False
          elif ((STATE == 17) and not EXT_CtrlCmd[EXT_ADDRESS_CMD_ABORT]):
              CMD_Abort = False
          end
          # ---------- Stop ---------- #
          if ((not STATE == 1) and (not STATE == 2) and (get_standard_digital_in(IO_ADDRESS_CMD_STOP) or EXT_CtrlCmd[EXT_ADDRESS_CMD_STOP])):
              CMD_Stop = True
              if get_standard_digital_in(IO_ADDRESS_CMD_STOP):
                  log_state("Stop command by pushbutton")
              elif EXT_CtrlCmd[EXT_ADDRESS_CMD_STOP]:
                  log_state("Stop command by external control")
              end
          elif (STATE == 2) and (not get_standard_digital_in(IO_ADDRESS_CMD_STOP)) and (not EXT_CtrlCmd[EXT_ADDRESS_CMD_STOP]):
              CMD_Stop = False
          end
          CMD_Hold = (STATE == 6 or STATE == 10) and not CMD_Stop and (ERROR.FLAG or EXT_CtrlCmd[EXT_ADDRESS_CMD_HOLD])
          CMD_Reset = (STATE == 2 or STATE == 8) and not CMD_Stop and (read_input_boolean_register(5) or EXT_CtrlCmd[EXT_ADDRESS_CMD_RESET])
          CMD_Start = (STATE == 4) and not CMD_Stop and (get_standard_digital_in(IO_ADDRESS_CMD_START) or EXT_CtrlCmd[EXT_ADDRESS_CMD_START])
          CMD_Unhold = (STATE == 10) and not CMD_Stop and (get_standard_digital_in(IO_ADDRESS_CMD_START) or EXT_CtrlCmd[EXT_ADDRESS_CMD_UNHOLD])
          CMD_Suspend = (STATE == 6) and not CMD_Stop and (CND_Suspend or EXT_CtrlCmd[EXT_ADDRESS_CMD_SUSPEND])
          CMD_Unsuspend = (STATE == 13) and not CMD_Stop and (CND_Unsuspend or EXT_CtrlCmd[EXT_ADDRESS_CMD_UNSUSPEND])
          CMD_Clear = (STATE == 16) and EXT_CtrlCmd[EXT_ADDRESS_CMD_CLEAR]
          FNC_Freedrive = (STATE == 10) and EXT_CtrlCmd[EXT_ADDRESS_FNC_FREEDRIVE]
          sleep(0.1)
      end
  end

  thread_pml_command_handler = run Get_Pml_Command()

  def command_manager(external_control="uGO", cond_suspend=False, cond_unsuspend=False):

      EXT_Control_by = external_control
      CND_Suspend = cond_suspend
      CND_Unsuspend = cond_unsuspend

      if (CMD_Abort and STATE != 15 and STATE != 16):
          STATE = 15
      elif (CMD_Stop and STATE != 1 and STATE != 2):
          STATE = 1
      end
      return False
  end

  def stopping():
      if (EXT_Control_by == "uGO"):
          return ugo_pml_stopping()
      elif (EXT_Control_by == "Leitsystem"):
          # EXT_CtrlCmd = Leitsystem
      else:
          return True
      end
      return False
  end

  def resetting():
      if (EXT_Control_by == "uGO"):
          return ugo_pml_resetting()
      elif (EXT_Control_by == "Leitsystem"):
          # EXT_CtrlCmd = Leitsystem
      else:
          return True
      end
      return False
  end

  def starting():
      if (EXT_Control_by == "uGO"):
          return ugo_pml_starting()
      elif (EXT_Control_by == "Leitsystem"):
          # EXT_CtrlCmd = Leitsystem
      else:
          return True
      end
      return False
  end

  def holding():
      if (EXT_Control_by == "uGO"):
          return ugo_pml_holding()
      elif (EXT_Control_by == "Leitsystem"):
          # EXT_CtrlCmd = Leitsystem
      else:
          return True
      end
      return False
  end

  def unholding():
      if (EXT_Control_by == "uGO"):
          return ugo_pml_unholding()
      elif (EXT_Control_by == "Leitsystem"):
          # EXT_CtrlCmd = Leitsystem
      else:
          return True
      end
      return False
  end

  def suspending():
      if (EXT_Control_by == "uGO"):
          return ugo_pml_suspending()
      elif (EXT_Control_by == "Leitsystem"):
          # EXT_CtrlCmd = Leitsystem
      else:
          return True
      end
      return False
  end

  def unsuspending():
      if (EXT_Control_by == "uGO"):
          return ugo_pml_unsuspending()
      elif (EXT_Control_by == "Leitsystem"):
          # EXT_CtrlCmd = Leitsystem
      else:
          return True
      end
      return False
  end

  def completing():
      if (EXT_Control_by == "uGO"):
          return ugo_pml_completing()
      elif (EXT_Control_by == "Leitsystem"):
          # EXT_CtrlCmd = Leitsystem
      else:
          return True
      end
      return False
  end

  def aborting():
      if (EXT_Control_by == "uGO"):
          return ugo_pml_aborting()
      elif (EXT_Control_by == "Leitsystem"):
          # EXT_CtrlCmd = Leitsystem
      else:
          return True
      end
      return False
  end

  def clearing():
      if (EXT_Control_by == "uGO"):
          return ugo_pml_clearing()
      elif (EXT_Control_by == "Leitsystem"):
          # EXT_CtrlCmd = Leitsystem
      else:
          return True
      end
      return False
  end
  $ 8 "Script: SCRIPT Utility V5.5.script"
  #*****************************************************
  # customer          :   tbd
  # project name      :   tbd
  #****************************************************
  # controller        :
  # software          :
  #****************************************************
  # author            :   P. Koehnke (+49 1628859904; p.koehnke@unitedrobotics.group)
  # Copyright (c)     :   United Robotics Group Health and Food GmbH
  #                       An der Riede 2
  #                       28816 Stuhr
  #                       Germany
  #****************************************************
  # description       :   utility programs for the application
  # version:      	:   3.1
  # created           :   30.01.2023
  # updated           :
  #****************************************************
  # modifications     :   get_tool_free_pose_2(), get_index_from_list()
  #
  # date              :   05.01.2024
  # name              :   PK
  # reason            :
  #****************************************************

  def found_in_matrix(data, req_id, req_idx):
      local id = -1
      local dimensions = size(data)
      local loop_dataset = 0

      while (id != req_id and loop_dataset < dimensions[0]):
          id = data[loop_dataset, 0]
          if (id == req_id):
              return data[loop_dataset, req_idx]
          else:
              loop_dataset = loop_dataset + 1
          end
      end
  end

  def found_in_list(value, list):
      local idx = 0

      while (idx < length(list)):
          if (value == list[idx]):
              return True
          end
          idx = idx + 1
      end
      return False
  end

  def get_index_from_list(list, value = -1):
      local idx = 0

      while (idx < length(list)):
          if (value == -1):
              if (list[idx] != 0):
                  return idx
              end
          else:
              if (list[idx] == value):
                  return idx
              end
          end
          idx = idx + 1
      end
      return -1
  end

  def find_object_by_type(list, type=0):
      local object = list[0]
      local i = 0

      while i < length(list):
          object = list[i]
          if object.type == type:
              return object
          end
          i = i + 1
      end
  end

  def pose_RPY2RotVec(pose):
      local rotvec = rpy2rotvec([d2r(pose[3]), d2r(pose[4]), d2r(pose[5])])
      return p[pose[0], pose[1], pose[2], rotvec[0], rotvec[1], rotvec[2]]
  end

  def pose_RotVec2RPY(pose):
      local rpy = rotvec2rpy([pose[3], pose[4], pose[5]])
      return p[pose[0], pose[1], pose[2], r2d(rpy[0]), r2d(rpy[1]), r2d(rpy[2])]
  end

  def swivel(frame_ref, angles = [0, 0, 0], pose = p[0, 0, 0, 0, 0, 0]):

      local rpy_ref = [0, 0, 0]
      local rpy_new = [0, 0, 0]
      local rotvec_new = [0, 0, 0]
      local pose_from = p[0, 0, 0, 0, 0, 0]
      local pose_to = p[0, 0, 0, 0, 0, 0]
      local i = 0

      if (pose == p[0, 0, 0, 0, 0, 0]):
          pose_to = pose_trans(pose_inv(frame_ref), get_actual_tcp_pose())
      else:
          pose_to = pose
      end

      rpy_ref = rotvec2rpy(frame_ref[3], frame_ref[4], frame_ref[5])

      while (i < 3):
          rpy_new[i] = rpy_ref[i] + d2r(angles[i])
          i = i + 1
      end

      rotvec_new = rpy2rotvec(rpy_new)
      pose_from = p[0, 0, 0, rotvec_new[0], rotvec_new[1], rotvec_new[2]]
      pose_to = p[pose_to[0], pose_to[1], pose_to[2], rotvec_new[0], rotvec_new[1], rotvec_new[2]]

      return pose_trans(pose_from, pose_to)
  end

  def get_random_pose(pose_ref, mode = "", range_max = [0, 0, 0]):
      # modi: "cubic", "rotation"
      # getting a random pose in the x/y-plane. range can be set for each
      # translation and rotation.
      local rpy_random = [0, 0, 0]
      local rotvec_random = [0, 0, 0]
      local pose_random = pose_ref
      local i = 0

      if (mode == "cubic"):
          # cubic mode: random pose takes only x, y and z
          i = 0
          while (i < 3):
              pose_random[i] = pose_ref[i] + range_max[i] * (random() - 0.5)
              i = i + 1
          end
          return pose_random

      elif (mode == "rotation"):
          i = 0
          while (i < 3):
              rpy_random[i] = d2r(range_max[i]) * (random() - 0.5)
              i = i + 1
          end
          rotvec_random = rpy2rotvec(rpy_random)
          pose_random = pose_trans(p[0, 0, 0, rotvec_random[0], rotvec_random[1], rotvec_random[2]], pose_ref)
          return pose_random

      else:
          # unknown mode, return pose_ref
          return pose_ref
      end
  end

  def get_pattern_pos_rectangle(counter, direction, pattern, patterninc = [0, 0], patternsize = [0, 0]):
      # defines the position inside a rectangular pattern
      # pattern describes, how many objects are in x-direction and how many in y-direction [x, y]
      # patternsize will give the total length of each direction [x, y]
      local X_Fac = 0
      local Y_Fac = 0
      local max = pattern[0] * pattern[1]
      local i = 0

      if (1 > counter or counter > max):
          counter = 1
      end

      if pattern[0] == 0:
          pattern[0] = 1
      end

      if pattern[1] == 0:
          pattern[1] = 1
      end

      if (direction == "Y" or direction == "y"):
          X_Fac = floor((counter - 1) / pattern[1])
          Y_Fac = (counter - 1) % pattern[1]
      elif (direction == "X" or direction == "x"):
          X_Fac = (counter - 1) % pattern[0]
          Y_Fac = floor((counter - 1) / pattern[0])
      end

      if patternsize != [0, 0]:
          while i < 2:
              if pattern[i] > 1:
                  patterninc[i] = patternsize[i] / (pattern[i] - 1)
              end
              i = i + 1
          end
      end

      return p[X_Fac * patterninc[0], Y_Fac * patterninc[1], 0, 0, 0, 0]
  end

  def get_pattern_pos_circle(counter, radius, angle, direction, pattern, patternsize = [0, 0]):
      # get the patternpos for a circular pattern through a counter
      # need the radius and the angle in radiants
      local X_Fac = 0
      local Y_Fac = 0
      local rad_bow = 0
      local radius_cal = 0
      local ref = p[0, 0, 0, 0, 0, 0]

      if pattern[0] == 0:
          pattern[0] = 1
      end

      if pattern[1] == 0:
          pattern[1] = 1
      end

      if (direction == "Y" or direction == "y"):
          X_Fac = floor((counter - 1) / pattern[1])
          Y_Fac = (counter - 1) % pattern[1]
      elif (direction == "X" or direction == "x"):
          X_Fac = (counter - 1) % pattern[0]
          Y_Fac = floor((counter - 1) / pattern[0])
      end

      # the opening angle will be calculated in x-direction
      # works only between -90 and 90 degree
      if pattern[0] > 1:
          rad_bow = - angle / (pattern[0] - 1) * X_Fac + angle / 2
      end

      if (counter % 2 == 0 and pattern[1] > 1):
          radius_cal = radius - patternsize[1] / (pattern[1])
      else:
          radius_cal = radius + patternsize[1] / (pattern[1])
      end
      ref = p[0, radius_cal, 0, 0, 0, 0]

      return p[ref[0] * cos(rad_bow) - ref[1] * sin(rad_bow), (ref[0] * sin(rad_bow) + ref[1] * cos(rad_bow)) - radius, 0, 0, 0, 0]
  end

  def get_pattern_counter(pose, direction, pattern, patterninc = [0, 0], patternsize = [0, 0]):
      # returns the counter for a pattern from a given cartesian pose
      local patternpose = p[pose[0], pose[1], 0, 0, 0, 0]
      local X_Fac = 0
      local Y_Fac = 0
      local i = 0

      if patternsize != [0, 0]:
          while i < 2:
              if pattern[i] > 1:
                  patterninc[i] = patternsize[i] / (pattern[i] - 1)
              else:
                  pattern[i] = 0
              end
              i = i + 1
          end
      end

      # calculation of the counter in the desired axis-direction
      if (direction == "x" or direction == "X"):
          if patterninc[0] > 0:
              X_Fac = ceil((patternpose[0] + patterninc[0] / 2) / patterninc[0])
              if X_Fac < 0:
                  X_Fac = 0
              end
          end
          if patterninc[1] > 0:
              Y_Fac = floor((patternpose[1] + patterninc[1] / 2) / patterninc[1])
              if Y_Fac < 0:
                  Y_Fac = 0
            end
          end
          return Y_Fac * pattern[0] + X_Fac
      elif (direction == "y" or direction == "Y"):
          if patterninc[0] > 0:
              X_Fac = floor((patternpose[0] + patterninc[0] / 2) / patterninc[0])
          end
          if patterninc[1] > 0:
              Y_Fac = ceil((patternpose[1] + patterninc[1] / 2) / patterninc[1])
          end
          return X_Fac * pattern[1] + Y_Fac
      end
  end

  def get_plc_reg(mod_sig_name):
      return integer_to_binary_list(modbus_get_signal_status(mod_sig_name))
  end

  def set_plc_reg(mod_sig_name, mod_sig_list):
      modbus_set_output_register(mod_sig_name, binary_list_to_integer(mod_sig_list), False)
  end

  def check_decapping(offset = 0, timeout = 5, abort = False):
      # checken, ob der Deckel schon ab ist
      local start = get_actual_tcp_pose()
      local current_offset = 0
      local timecounter = 0
      while (current_offset < offset and not abort):
          current_offset = pose_dist(start, get_actual_tcp_pose())
          timecounter = timecounter + 1
          if (timecounter * 0.5 == timeout):
              break
          end
          sleep(0.5)
      end
      stopl(0.5)
  end

  def check_capping(torque = 0):
      # checken, wann der Deckel verschraubt ist
      force_mode(get_actual_tcp_pose(), [0, 0, 1, 0, 0, 0], [0, 0, -2.0, 0, 0, 0], 2, [0.01, 0.01, 0.001, 0.01, 0.01, 0.01])
  end

  def is_reachable(frame, poses, offsets = [0, 0, 0]):
      local idx = 0
      local pose = p[0, 0, 0, 0, 0, 0]

      while (idx < length(poses)):
          pose = poses[idx]
          pose[0] = pose[0] + offsets[0]
          pose[1] = pose[1] + offsets[1]
          pose[2] = pose[2] + offsets[2]

          if pose != p[0, 0, 0, 0, 0, 0]:
              if (not get_inverse_kin_has_solution(pose_trans(frame, pose))):
                  textmsg(str_cat(str_cat("Pose ", to_str(idx + 1)), " is not reachable"))
                  return False
              end
          end
          idx = idx + 1
      end
      return True
  end

  def is_within_limits(frame, poses, offsets = [0, 0, 0]):
      local idx = 0
      local pose = p[0, 0, 0, 0, 0, 0]

      while (idx < length(poses)):
          pose = poses[idx]
          pose[0] = pose[0] + offsets[0]
          pose[1] = pose[1] + offsets[1]
          pose[2] = pose[2] + offsets[2]

          if is_reachable(frame = frame, poses = poses, offsets = offsets):
              if (not is_within_safety_limits(get_inverse_kin(pose_trans(frame, pose), get_actual_joint_positions()))):
                  textmsg(str_cat(str_cat("Pose ", to_str(idx + 1)), "is out of joint limits"))
                  return False
              else:
                  idx = idx + 1
              end
          else:
              return False
          end
      end
      return True
  end


  def string_to_list(string, separator = "," , endDelimiter = ";" , capacity = 50):
      local string_length = str_len(string)
      local list_out = make_list(length = elements_in_string(string), initial_value = -1, capacity = capacity)
      local cnt = 0
      local idx = 0

      while cnt < string_length-1 :
        textmsg("new loop")
        textmsg(to_str(idx))
        local sepAt = str_find(string, separator, cnt)
        textmsg(to_str(sepAt))
        if sepAt < 0 :
            sepAt = str_find(string, endDelimiter, cnt)
        end
        list_out[idx] = to_num(str_sub(string, cnt, sepAt-cnt))
        idx = idx +1
        cnt = sepAt + 1
      end

      return list_out
  end

  def elements_in_string(string, separator = "," , endDelimiter = ";" , capacity = 50):
     local string_length = str_len(string)
      local len = 0
      local sepAt = 0

      while sepAt < string_length-1 and sepAt>=0 :
        local sepAt = str_find(string, separator, sepAt+1)
        len = len +1
      end

      return len
  end
  $ 9 "Script: SCRIPT uML Lights V1.2.script"

  #****************************************************
  # product           : uLabMobile
  # language          : urscript
  #****************************************************
  # author            :   D.Kreugel
  # Copyright (c)     :   United Robotics Group
  #                       An der Riede 2
  #                       28816 Stuhr
  #                       Germany
  #****************************************************
  # description       :   led controls for uLabMobile
  # version:      	:   1.2
  # created           :   09.08.2024
  # updated           :
  #****************************************************
  # modifications     :   changed conditions to switch lights (not only pml state but also charging state)
  #
  # date              :   09.08.2024
  # name              :   PK
  # reason            :   due to the change in project P1117, we run to often through every state. This leads to to much colorchanges
  #****************************************************

  # HARDWARE CONFIGURATION
  LED_GREEN = struct(type="CO",id=5)
  LED_RED = struct(type="CO",id=6)
  LED_BLUE = struct(type="CO",id=7)

  def set_output(type,id,state=True):
      if(type=="CO"):
          set_configurable_digital_out(id,state)
      elif(type=="DO"):
          set_standard_digital_out(id,state)
      end
  end

  def led_red_on():
      set_output(LED_RED.type,LED_RED.id,True)
  end

  def led_red_off():
      set_output(LED_RED.type,LED_RED.id,False)
  end

  def led_green_on():
      set_output(LED_GREEN.type,LED_GREEN.id,True)
  end

  def led_green_off():
      set_output(LED_GREEN.type,LED_GREEN.id,False)
  end

  def led_blue_on():
      set_output(LED_BLUE.type,LED_BLUE.id,True)
  end

  def led_blue_off():
      set_output(LED_BLUE.type,LED_BLUE.id,False)
  end


  # COLOR MIX
  def color_blue():
      led_blue_on()
      led_green_off()
      led_red_off()
  end

  def color_red():
      led_blue_off()
      led_green_off()
      led_red_on()
  end

  def color_green():
      led_blue_off()
      led_green_on()
      led_red_off()
  end

  def color_yellow():
      led_blue_off()
      led_green_on()
      led_red_on()
  end

  def color_lightblue():
      led_blue_on()
      led_green_on()
      led_red_off()
  end

  def color_violet():
      led_blue_on()
      led_green_off()
      led_red_on()
  end

  def color_white():
      led_blue_on()
      led_green_on()
      led_red_on()
  end

  def led_off():
      led_blue_off()
      led_green_off()
      led_red_off()
  end

